      rq_wait_pos_spe_for_request(255, 204, 255, "1")
      rq_go_to("1")
      rq_wait("1")
      # end: URCap Program Node
      $ 2057 "Decap"
      $ 2058 "Action_Info≔'decapping'"
      global Action_Info="decapping"
      $ 2059 "Set GRP_3F_Enable=On"
      set_standard_digital_out(4, True)
      $ 2060 "Set GRP_3F_Decap=On"
      set_standard_digital_out(3, True)
      $ 2061 "Force"
      sleep(0.02)
      zero_ftsensor()
      force_mode(p[0.0,0.0,0.0,0.0,0.0,0.0], [0, 0, 1, 0, 0, 0], [0.0, 0.0, 1.0, 0.0, 0.0, 0.0], 2, [0.1, 0.1, 0.001, 0.3490658503988659, 0.3490658503988659, 0.3490658503988659])
      $ 2062 "check_decapping(offset=0.015, timeout=10, abort=CMD_Hold)" "noBreak"
      check_decapping(offset=0.015, timeout=10, abort=CMD_Hold)
      end_force_mode()
      stopl(5.0)
      $ 2063 "Set GRP_3F_Decap=Off"
      set_standard_digital_out(3, False)
      $ 2064 "Set GRP_3F_Enable=Off"
      set_standard_digital_out(4, False)
      $ 2065 "MoveL"
      $ 2066 "Waypoint_90" "breakAfter"
      movel(Waypoint_90_p, a=0.5, v=0.1, r=0.05)
      $ 2067 "MoveJ"
      $ 2068 "cap_dump_2" "breakAfter"
      movej(get_inverse_kin(cap_dump_2_p, qnear=cap_dump_2_q), a=0.5235987755982988, v=0.4363323129985824)
      # begin: URCap Program Node
      #   Source: Robotiq_Grippers, 3.17.0.105337, Robotiq Inc.
      #   Type: Gripper
      $ 2069 "Gripper Open (1)"
      if not(gripper_connected[0]):
        popup("Gripper 1 must be connected to run this program.", "No connection", False, True, True)
      end
      if not(rq_is_gripper_activated("1")):
        popup("Gripper 1 is not activated. Go to Installation tab > Gripper to activate it and run the program again.", "Not activated", False, True, True)
      end
      rq_set_pos_spd_for(0, 204, 255, "1")
      rq_wait_pos_spe_for_request(0, 204, 255, "1")
      rq_go_to("1")
      rq_wait("1")
      # end: URCap Program Node
      $ 2070 "MoveJ"
      $ 2071 "Waypoint_91" "breakAfter"
      movej(get_inverse_kin(Waypoint_91_p, qnear=Waypoint_91_q), a=0.5235987755982988, v=0.4363323129985824, r=0.036)
    elif (33 == switch_1):
      $ 2072 "Case 33"
      $ 2073 "Shake and liquid transfer"
      $ 2074 "MoveL"
      $ 2075 "Vial_liq_abov_1" "breakAfter"
      movel(Vial_liq_abov_1_p, a=0.5, v=0.1)
      $ 2076 "Vial_liq_pick_3" "breakAfter"
      movel(Vial_liq_pick_3_p, a=0.5, v=0.1)
      $ 2077 "Vial_liq_pick_4" "breakAfter"
      movel(Vial_liq_pick_4_p, a=0.5, v=0.1)
      # begin: URCap Program Node
      #   Source: Robotiq_Grippers, 3.17.0.105337, Robotiq Inc.
      #   Type: Gripper
      $ 2078 "Gripper Close (1)"
      if not(gripper_connected[0]):
        popup("Gripper 1 must be connected to run this program.", "No connection", False, True, True)
      end
      if not(rq_is_gripper_activated("1")):
        popup("Gripper 1 is not activated. Go to Installation tab > Gripper to activate it and run the program again.", "Not activated", False, True, True)
      end
      rq_set_pos_spd_for(255, 82, 71, "1")
      rq_wait_pos_spe_for_request(255, 82, 71, "1")
      rq_go_to("1")
      rq_wait("1")
      # end: URCap Program Node
      $ 2079 "Wait: 1.0"
      sleep(1.0)
      $ 2080 "Set GRP_3F_Open=On"
      set_standard_digital_out(5, True)
      $ 2081 "Wait: 0.5"
      sleep(0.5)
      $ 2082 "Vial_liq_abov_2" "breakAfter"
      movel(Vial_liq_abov_2_p, a=0.3, v=0.05, r=0.05)
      $ 2083 "MoveL"
      $ 2084 "Liquid_midway_1" "breakAfter"
      movel(Liquid_midway_1_p, a=0.5, v=0.1)
      $ 2085 "Loop 3 times"
      Loop_1 = 0
      while (Loop_1 < 3):
        $ 2086 "shake_3" "breakAfter"
        movel(shake_3_p, a=2.0, v=0.5)
        $ 2087 "shake_4" "breakAfter"
        movel(shake_4_p, a=2.0, v=0.5)
        Loop_1 = Loop_1 + 1
      end
      $ 2088 "drop_above_3" "breakAfter"
      movel(drop_above_3_p, a=0.5, v=0.1)
      $ 2089 "drop_above_4" "breakAfter"
      movel(drop_above_4_p, a=0.5, v=0.1)
      $ 2090 "liq_tran_3" "breakAfter"
      movel(liq_tran_3_p, a=0.5, v=0.05, r=0.008)
      $ 2091 "Wait: 1.0"
      sleep(1.0)
      $ 2092 "drop_above_5" "breakAfter"
      movel(drop_above_5_p, a=0.5, v=0.1)
      $ 2093 "Waypoint_92" "breakAfter"
      movel(Waypoint_92_p, a=0.5, v=0.1)
      $ 2094 "liq_tran_4" "breakAfter"
      movel(liq_tran_4_p, a=0.5, v=0.05)
      $ 2095 "Wait: 1.0"
      sleep(1.0)
      $ 2096 "drop_above_6" "breakAfter"
      movel(drop_above_6_p, a=0.5, v=0.1)
      $ 2097 "drop_above_7" "breakAfter"
      movel(drop_above_7_p, a=0.5, v=0.1)
      $ 2098 "Liquid_midway_2" "breakAfter"
      movel(Liquid_midway_2_p, a=0.5, v=0.1)
      $ 2099 "MoveL"
      $ 2100 "Vial_drop_abo_1" "breakAfter"
      movel(Vial_drop_abo_1_p, a=0.5, v=0.1)
      $ 2101 "Vial_liq_drop_1" "breakAfter"
      movel(Vial_liq_drop_1_p, a=0.5, v=0.1)
      # begin: URCap Program Node
      #   Source: Robotiq_Grippers, 3.17.0.105337, Robotiq Inc.
      #   Type: Gripper
      $ 2102 "Gripper Open (1)"
      if not(gripper_connected[0]):
        popup("Gripper 1 must be connected to run this program.", "No connection", False, True, True)
      end
      if not(rq_is_gripper_activated("1")):
        popup("Gripper 1 is not activated. Go to Installation tab > Gripper to activate it and run the program again.", "Not activated", False, True, True)
      end
      rq_set_pos_spd_for(0, 82, 71, "1")
      rq_wait_pos_spe_for_request(0, 82, 71, "1")
      rq_go_to("1")
      rq_wait("1")
      # end: URCap Program Node
      $ 2103 "Vial_drop_abo_2" "breakAfter"
      movel(Vial_drop_abo_2_p, a=0.5, v=0.1)
    elif (34 == switch_1):
      $ 2104 "Case 34"
      $ 2105 "Task≔'Dosing'"
      global Task="Dosing"
      $ 2106 "tilt_to_home()"
      tilt_to_home()
      $ 2107 "Powder dosing all"
      $ 2108 "tilt_angle_sent≔0.0"
      global tilt_angle_sent=0.0
      $ 2109 "send_target_info()"
      send_target_info()
      $ 2111 "prev_spat≔''"
      global prev_spat=""
      $ 2112 "spatula≔''"
      global spatula=""
      $ 2113 "scoop_status≔'normal'"
      global scoop_status="normal"
      $ 2114 "send_powder_info()"
      send_powder_info()
      $ 2115 "Set AO[0]=0.0"
      set_standard_analog_out(0, 0.0)
      $ 2116 "Wait: 0.2"
      sleep(0.2)
      $ 2117 "reach pots decapping pose"
      # begin: URCap Program Node
      #   Source: SensoPart VISOR Robotic, 2.0.6, SensoPart Industriesensorik GmbH
      #   Type: VISOR Robotic App
      $ 2123 "VISOR Easy Pick"
      def visorFuncEasyPick_4c19ec():
        # begin: URCap Program Node
        #   Source: SensoPart VISOR Robotic, 2.0.6, SensoPart Industriesensorik GmbH
        #   Type: Easy Pick Setup
        $ 2124 "# 1 Setup" "noBreak"
        local easyPickVisorId = 1
        local easyPickArmMounted = True
        local easyPickSetJob = True
        local easyPickJobName = "Weight_scale"
        local easyPickAtImgAcq = False
        local easyPickImgAcqPose = Trigger
        # end: URCap Program Node
        # begin: URCap Program Node
        #   Source: SensoPart VISOR Robotic, 2.0.6, SensoPart Industriesensorik GmbH
        #   Type: Process
        $ 2125 "Process" "noBreak"
        local easyPickObjTaken = False
        local easyPickTrigger = False
        local easyPickPoseIdx = 0
        local easyPickPose = p[0,0,0,0,0,0]
        def easyPickFuncTrigger(visorId, setJob, jobName, arm):
        if (setJob):
          visor_changeJob(visorId, jobName, 6000)
        end
        if (arm):
          visor_trigger(visorId, 6000, "arm")
        else:
          visor_trigger(visorId, 6000)
        end
        global easyPickParts_4=visor_partsFound(visorId)
        visor_easyPickUpdate(visorId, "parts", visor_partsFound(visorId))
        return visor_getPose3d(visorId, 0)
      end
      while (not easyPickObjTaken):
        easyPickTrigger = (easyPickCount_4 >= visor_partsFound(easyPickVisorId)) or (easyPickCount_4 > 9) or (not visor_easyPickCheckIdent("3d3650", easyPickVisorId))
        if (easyPickTrigger):
          easyPickCount_4 = 0
        end
        easyPickPoseIdx = easyPickCount_4
        easyPickPose = visor_getPose3d(easyPickVisorId, easyPickPoseIdx)
        visor_easyPickUpdate(easyPickVisorId, "counter", easyPickPoseIdx)
        # begin: URCap Program Node
        #   Source: SensoPart VISOR Robotic, 2.0.6, SensoPart Industriesensorik GmbH
        #   Type: Image Acquisition Pose
        $ 2126 "Image Acquisition Pose" "noBreak"
        if (easyPickTrigger):
          if (not easyPickAtImgAcq):
            movej(pose_trans(easyPickImgAcqPose,p[0.0000,0.0000,-0.0000,0.0000,0.0000,0.0000]),a=1.3963,v=1.0472,t=0.000000,r=0.000000)
            easyPickAtImgAcq = True
          end
          easyPickPose = easyPickFuncTrigger(easyPickVisorId, easyPickSetJob, easyPickJobName, easyPickArmMounted)
        end
        # end: URCap Program Node
        # begin: URCap Program Node
        #   Source: SensoPart VISOR Robotic, 2.0.6, SensoPart Industriesensorik GmbH
        #   Type: Object Detected
        $ 2127 "Object Detected" "noBreak"
        if (visor_partsFound(easyPickVisorId) > 0):
          $ 2128 "Open Gripper" "noBreak"
          $ 2129 "weight_value≔get_weight()" "noBreak"
          global weight_value=get_weight()
          $ 2130 "Wait: 0.5" "noBreak"
          sleep(0.5)
          $ 2131 "diff≔target_weight-weight_value" "noBreak"
          global diff=target_weight-weight_value
          $ 2132 "compute_level_percent(W_now, weight_value)" "noBreak"
          compute_level_percent(W_now, weight_value)
          $ 2133 "send_level_info()" "noBreak"
          send_level_info()
          $ 2134 "spatula≔select_spatula(Flowability, level, diff, bulk_density, mouth_d)" "noBreak"
          global spatula=select_spatula(Flowability, level, diff, bulk_density, mouth_d)
          $ 2135 "Wait: 0.2" "noBreak"
          sleep(0.2)
          $ 2136 "send_spatula_info()" "noBreak"
          send_spatula_info()
          $ 2137 "Pick spatula" "noBreak"
          $ 2138 "If spatula ≟ 'spatula_L'" "noBreak"
          if (spatula  ==  "spatula_L"):
            $ 2139 "MoveJ" "noBreak"
            $ 2140 "Spatula_otw" "noBreak"
            movej(get_inverse_kin(Spatula_otw_p, qnear=Spatula_otw_q), a=1.3962634015954636, v=1.0471975511965976)
            $ 2141 "pick_spat_L_abv" "noBreak"
            movej(get_inverse_kin(pick_spat_L_abv_p, qnear=pick_spat_L_abv_q), a=1.3962634015954636, v=1.0471975511965976)
            $ 2142 "MoveL" "noBreak"
            $ 2143 "spat_L_pick" "noBreak"
            movel(spat_L_pick_p, a=1.2, v=0.25)
            # begin: URCap Program Node
            #   Source: Robotiq_Grippers, 3.17.0.105337, Robotiq Inc.
            #   Type: Gripper
            $ 2144 "Gripper Close (1)" "noBreak"
            if not(gripper_connected[0]):
              popup("Gripper 1 must be connected to run this program.", "No connection", False, True, True)
            end
            if not(rq_is_gripper_activated("1")):
              popup("Gripper 1 is not activated. Go to Installation tab > Gripper to activate it and run the program again.", "Not activated", False, True, True)
            end
            rq_set_pos_spd_for(255, 0, 77, "1")
            rq_wait_pos_spe_for_request(255, 0, 77, "1")
            rq_go_to("1")
            rq_wait("1")
            # end: URCap Program Node
            $ 2145 "spat_L_lift" "noBreak"
            movel(spat_L_lift_p, a=1.2, v=0.25, r=0.01)
            $ 2146 "spat_L_side" "noBreak"
            movel(spat_L_side_p, a=1.2, v=0.25, r=0.01)
            $ 2147 "spat_L_up" "noBreak"
            movel(spat_L_up_p, a=1.2, v=0.25, r=0.05)
            $ 2148 "MoveJ" "noBreak"
            $ 2149 "Spatula_otw" "noBreak"
            movej(get_inverse_kin(Spatula_otw_p, qnear=Spatula_otw_q), a=1.3962634015954636, v=1.0471975511965976)
          else:
            $ 2150 "ElseIf spatula ≟'spatula_M'" "noBreak"
            if (spatula  == "spatula_M"):
              $ 2151 "MoveJ" "noBreak"
              $ 2152 "Spatula_otw" "noBreak"
              movej(get_inverse_kin(Spatula_otw_p, qnear=Spatula_otw_q), a=1.3962634015954636, v=1.0471975511965976)
              $ 2153 "spat_M_up" "noBreak"
              movej(get_inverse_kin(spat_M_up_p, qnear=spat_M_up_q), a=1.3962634015954636, v=1.0471975511965976, r=0.05)
              $ 2154 "MoveL" "noBreak"
              $ 2155 "spat_M_pick" "noBreak"
              movel(spat_M_pick_p, a=1.2, v=0.25)
              # begin: URCap Program Node
              #   Source: Robotiq_Grippers, 3.17.0.105337, Robotiq Inc.
              #   Type: Gripper
              $ 2156 "Gripper Close (1)" "noBreak"
              if not(gripper_connected[0]):
                popup("Gripper 1 must be connected to run this program.", "No connection", False, True, True)
              end
              if not(rq_is_gripper_activated("1")):
                popup("Gripper 1 is not activated. Go to Installation tab > Gripper to activate it and run the program again.", "Not activated", False, True, True)
              end
              rq_set_pos_spd_for(255, 0, 77, "1")
              rq_wait_pos_spe_for_request(255, 0, 77, "1")
              rq_go_to("1")
              rq_wait("1")
              # end: URCap Program Node
              $ 2157 "spat_M_up" "noBreak"
              movel(spat_M_up_p, a=1.2, v=0.25, r=0.05)
              $ 2158 "Spatula_otw" "noBreak"
              movel(Spatula_otw_p, a=1.2, v=0.25)
              $ 2159 "switch_spat_M≔ False " "noBreak"
              global switch_spat_M=  False
            else:
              $ 2160 "ElseIf spatula≟'spatula_S'" "noBreak"
              if (spatula == "spatula_S"):
                $ 2161 "MoveJ" "noBreak"
                $ 2162 "Spatula_otw" "noBreak"
                movej(get_inverse_kin(Spatula_otw_p, qnear=Spatula_otw_q), a=1.3962634015954636, v=1.0471975511965976)
                $ 2163 "spat_S_Up_7" "noBreak"
                movej(get_inverse_kin(spat_S_Up_7_p, qnear=spat_S_Up_7_q), a=1.3962634015954636, v=1.0471975511965976, r=0.05)
                $ 2164 "MoveL" "noBreak"
                $ 2165 "spat_S_Pick_4" "noBreak"
                movel(spat_S_Pick_4_p, a=1.2, v=0.25)
                # begin: URCap Program Node
                #   Source: Robotiq_Grippers, 3.17.0.105337, Robotiq Inc.
                #   Type: Gripper
                $ 2166 "Gripper Close (1)" "noBreak"
                if not(gripper_connected[0]):
                  popup("Gripper 1 must be connected to run this program.", "No connection", False, True, True)
                end
                if not(rq_is_gripper_activated("1")):
                  popup("Gripper 1 is not activated. Go to Installation tab > Gripper to activate it and run the program again.", "Not activated", False, True, True)
                end
                rq_set_pos_spd_for(255, 0, 77, "1")
                rq_wait_pos_spe_for_request(255, 0, 77, "1")
                rq_go_to("1")
                rq_wait("1")
                # end: URCap Program Node
                $ 2167 "spat_S_Up_8" "noBreak"
                movel(spat_S_Up_8_p, a=1.2, v=0.25, r=0.05)
                $ 2168 "Spatula_otw" "noBreak"
                movel(Spatula_otw_p, a=1.2, v=0.25)
                $ 2169 "switch_spat_S≔ False " "noBreak"
                global switch_spat_S=  False
              else:
                $ 2170 "ElseIf spatula≟'spatula_flat_M'" "noBreak"
                if (spatula == "spatula_flat_M"):
                  $ 2171 "MoveJ" "noBreak"
                  $ 2172 "Spatula_otw" "noBreak"
                  movej(get_inverse_kin(Spatula_otw_p, qnear=Spatula_otw_q), a=1.3962634015954636, v=1.0471975511965976)
                  $ 2173 "spat_flatM_up" "noBreak"
                  movej(get_inverse_kin(spat_flatM_up_p, qnear=spat_flatM_up_q), a=1.3962634015954636, v=1.0471975511965976, r=0.05)
                  $ 2174 "MoveL" "noBreak"
                  $ 2175 "spat_flatM_pick" "noBreak"
                  movel(spat_flatM_pick_p, a=1.2, v=0.25)
                  # begin: URCap Program Node
                  #   Source: Robotiq_Grippers, 3.17.0.105337, Robotiq Inc.
                  #   Type: Gripper
                  $ 2176 "Gripper Close (1)" "noBreak"
                  if not(gripper_connected[0]):
                    popup("Gripper 1 must be connected to run this program.", "No connection", False, True, True)
                  end
                  if not(rq_is_gripper_activated("1")):
                    popup("Gripper 1 is not activated. Go to Installation tab > Gripper to activate it and run the program again.", "Not activated", False, True, True)
                  end
                  rq_set_pos_spd_for(255, 0, 77, "1")
                  rq_wait_pos_spe_for_request(255, 0, 77, "1")
                  rq_go_to("1")
                  rq_wait("1")
                  # end: URCap Program Node
                  $ 2177 "spat_flatM_up" "noBreak"
                  movel(spat_flatM_up_p, a=1.2, v=0.25, r=0.05)
                  $ 2178 "Spatula_otw" "noBreak"
                  movel(Spatula_otw_p, a=1.2, v=0.25)
                  $ 2179 "switch_spat_F_M≔ False " "noBreak"
                  global switch_spat_F_M=  False
                else:
                  $ 2180 "ElseIf spatula≟'spatula_flat_S'" "noBreak"
                  if (spatula == "spatula_flat_S"):
                    $ 2181 "MoveJ" "noBreak"
                    $ 2182 "Spatula_otw" "noBreak"
                    movej(get_inverse_kin(Spatula_otw_p, qnear=Spatula_otw_q), a=1.3962634015954636, v=1.0471975511965976)
                    $ 2183 "spat_flatS_up" "noBreak"
                    movej(get_inverse_kin(spat_flatS_up_p, qnear=spat_flatS_up_q), a=1.3962634015954636, v=1.0471975511965976, r=0.05)
                    $ 2184 "MoveL" "noBreak"
                    $ 2185 "spat_flatS_pick" "noBreak"
                    movel(spat_flatS_pick_p, a=1.2, v=0.25)
                    # begin: URCap Program Node
                    #   Source: Robotiq_Grippers, 3.17.0.105337, Robotiq Inc.
                    #   Type: Gripper
                    $ 2186 "Gripper Close (1)" "noBreak"
                    if not(gripper_connected[0]):
                      popup("Gripper 1 must be connected to run this program.", "No connection", False, True, True)
                    end
                    if not(rq_is_gripper_activated("1")):
                      popup("Gripper 1 is not activated. Go to Installation tab > Gripper to activate it and run the program again.", "Not activated", False, True, True)
                    end
                    rq_set_pos_spd_for(255, 0, 77, "1")
                    rq_wait_pos_spe_for_request(255, 0, 77, "1")
                    rq_go_to("1")
                    rq_wait("1")
                    # end: URCap Program Node
                    $ 2187 "spat_flatS_up" "noBreak"
                    movel(spat_flatS_up_p, a=1.2, v=0.25, r=0.05)
                    $ 2188 "Spatula_otw" "noBreak"
                    movel(Spatula_otw_p, a=1.2, v=0.25)
                    $ 2189 "switch_spat_F_S≔ False " "noBreak"
                    global switch_spat_F_S=  False
                  end
                end
              end
            end
          end
          $ 2190 "Action_Info≔'Scooping'" "noBreak"
          global Action_Info="Scooping"
          $ 2191 "auto_tilt_and_scoop(W_now, target_weight, weight_value)" "noBreak"
          auto_tilt_and_scoop(W_now, target_weight, weight_value)
          $ 2192 "Action_Info≔'Dosing'" "noBreak"
          global Action_Info="Dosing"
          # begin: URCap Program Node
          #   Source: SensoPart VISOR Robotic, 2.0.6, SensoPart Industriesensorik GmbH
          #   Type: Approach Pose
          $ 2193 "Approach Pose" "noBreak"
          movej(pose_trans(easyPickPose,p[0.0000,0.0000,-0.0000,0.0000,0.0000,0.0000]),a=0.2618,v=0.1745,t=0.000000,r=0.000000)
          # end: URCap Program Node
          # begin: URCap Program Node
          #   Source: SensoPart VISOR Robotic, 2.0.6, SensoPart Industriesensorik GmbH
          #   Type: Target Pose
          $ 2194 "Target Pose" "noBreak"
          movel(pose_trans(easyPickPose,p[0.0000,0.0000,-0.0000,0.0000,0.0000,0.0000]),a=0.0500,v=0.0200,t=0.000000,r=0.000000)
          # end: URCap Program Node
          $ 2195 "Close Gripper" "noBreak"
          $ 2196 "current_p≔get_actual_tcp_pose()" "noBreak"
          global current_p= get_actual_tcp_pose ()
          $ 2197 "dispense_pos≔pose_trans(current_p,p[0,0,0,0,-deg2rad(spatula_ry),0])" "noBreak"
          global dispense_pos=pose_trans(current_p,p[0,0,0,0,-deg2rad(spatula_ry),0])
          $ 2198 "Loop weight_value≤target_weight and delta_count≤3" "noBreak"
          thread Thread_while_2198():
            while (True):
              $ 2199 "MoveL" "noBreak"
              $ 2200 "dispense_pos" "noBreak"
              movel(dispense_pos, a=0.2, v=0.1)
              $ 2201 "log_weight()" "noBreak"
              log_weight()
              $ 2203 "CCW_full_Rotate()" "noBreak"
              CCW_full_Rotate()
              $ 2204 "Start_thread≔ True " "noBreak"
              global Start_thread=  True
              $ 2205 "vib_thread≔ True " "noBreak"
              global vib_thread=  True
              $ 2206 "Wait: 0.5" "noBreak"
              sleep(0.5)
              $ 2207 "If diff ≥(target_g*1.2)" "noBreak"
              if (diff  >= (target_g*1.2)):
                $ 2208 "tilt_pose≔pose_trans(get_actual_tcp_pose(), p[0, 0, 0, 0, 0, 2.0])" "noBreak"
                global tilt_pose=pose_trans(get_actual_tcp_pose(), p[0, 0, 0, 0, 0, 2.0])
                $ 2209 "movel(tilt_pose, a=0.5, v=0.5, r=0.00001)" "noBreak"
                movel(tilt_pose, a=0.5, v=0.5, r=0.00001)
              else:
                $ 2210 "Else" "noBreak"
                $ 2211 "Loop weight_value≤(target_weight-0.00) and tilt_angle≥(-1.999) and tilt_angle≤0.5" "noBreak"
                thread Thread_while_2211():
                  while (True):
                    $ 2212 "current_error≔target_weight-weight_value" "noBreak"
                    global current_error=target_weight-weight_value
                    $ 2213 "Integral_error≔Integral_error+current_error*dt" "noBreak"
                    global Integral_error=Integral_error+current_error*dt
                    $ 2214 "derivative≔(current_error-previous_error)/dt" "noBreak"
                    global derivative=(current_error-previous_error)/dt
                    $ 2215 "tilt_increment≔(kp*current_error)+(ki*Integral_error)+(kd*derivative)" "noBreak"
                    global tilt_increment=(kp*current_error)+(ki*Integral_error)+(kd*derivative)
                    $ 2216 "current_pose≔get_actual_tcp_pose()" "noBreak"
                    global current_pose= get_actual_tcp_pose ()
                    $ 2217 "tilt_angle≔current_pose[5]" "noBreak"
                    global tilt_angle=current_pose[5]
                    $ 2218 "tilt_pose≔pose_trans(current_pose, p[0, 0, 0, 0, 0, tilt_increment])" "noBreak"
                    global tilt_pose=pose_trans(current_pose, p[0, 0, 0, 0, 0, tilt_increment])
                    $ 2219 "movel(tilt_pose, a=0.1, v=0.1, r=0.00001)" "noBreak"
                    movel(tilt_pose, a=0.1, v=0.1, r=0.00001)
                    $ 2220 "previous_error≔current_error" "noBreak"
                    global previous_error=current_error
                  end
                end
                if (weight_value <= (target_weight-0.00)  and  tilt_angle >= (-1.999)  and  tilt_angle <= 0.5):
                  global thread_handler_2211=run Thread_while_2211()
                  while (weight_value <= (target_weight-0.00)  and  tilt_angle >= (-1.999)  and  tilt_angle <= 0.5):
                    sync()
                  end
                  kill thread_handler_2211
                end
              end
              $ 2221 "weight_value≔get_weight()" "noBreak"
              global weight_value=get_weight()
              $ 2222 "tilt_angle≔-1" "noBreak"
              global tilt_angle=-1
              $ 2223 "Wait: 0.5" "noBreak"
              sleep(0.5)
              $ 2224 "Start_thread≔ False " "noBreak"
              global Start_thread=  False
              $ 2225 "vib_thread≔ False " "noBreak"
              global vib_thread=  False
              $ 2226 "dispense_pos" "noBreak"
              movel(dispense_pos, a=1.2, v=0.25)
              $ 2227 "compute_level_percent(W_now, weight_value)" "noBreak"
              compute_level_percent(W_now, weight_value)
              $ 2228 "If delta<0.01" "noBreak"
              if (delta<0.01):
                $ 2229 "delta_count≔delta_count+1" "noBreak"
                global delta_count=delta_count+1
              else:
                $ 2230 "Else" "noBreak"
                $ 2231 "delta_count≔0" "noBreak"
                global delta_count=0
              end
              $ 2232 "prev_spat≔spatula" "noBreak"
              global prev_spat=spatula
              $ 2233 "Wait: 0.2" "noBreak"
              sleep(0.2)
              $ 2234 "spatula≔select_spatula(Flowability, level, diff, bulk_density, mouth_d)" "noBreak"
              global spatula=select_spatula(Flowability, level, diff, bulk_density, mouth_d)
              $ 2235 "Wait: 1.0" "noBreak"
              sleep(1.0)
              $ 2236 "send_level_info()" "noBreak"
              send_level_info()
              $ 2237 "send_spatula_info()" "noBreak"
              send_spatula_info()
              $ 2238 "Integral_error≔0" "noBreak"
              global Integral_error=0
              $ 2239 "current_error≔0" "noBreak"
              global current_error=0
              $ 2240 "previous_error≔0" "noBreak"
              global previous_error=0
              $ 2241 "Set AO[0]=0.0" "noBreak"
              set_standard_analog_out(0, 0.0)
              $ 2242 "Wait: 0.5" "noBreak"
              sleep(0.5)
              $ 2243 "swtich spatula" "noBreak"
              $ 2244 "If spatula ≟ 'spatula_M' and switch_spat_M≟ True " "noBreak"
              if (spatula  ==  "spatula_M"  and  switch_spat_M ==   True  ):
                $ 2245 "MoveJ" "noBreak"
                $ 2246 "Spatula_otw" "noBreak"
                movej(get_inverse_kin(Spatula_otw_p, qnear=Spatula_otw_q), a=1.3962634015954636, v=1.0471975511965976)
                $ 2247 "spat_L_up" "noBreak"
                movej(get_inverse_kin(spat_L_up_p, qnear=spat_L_up_q), a=1.3962634015954636, v=1.0471975511965976)
                $ 2248 "MoveL" "noBreak"
                $ 2249 "spat_L_side" "noBreak"
                movel(spat_L_side_p, a=1.2, v=0.25)
                $ 2250 "spat_L_lift" "noBreak"
                movel(spat_L_lift_p, a=1.2, v=0.25)
                $ 2251 "spat_L_pick" "noBreak"
                movel(spat_L_pick_p, a=0.2, v=0.1)
                # begin: URCap Program Node
                #   Source: Robotiq_Grippers, 3.17.0.105337, Robotiq Inc.
                #   Type: Gripper
                $ 2252 "Gripper Open (1)" "noBreak"
                if not(gripper_connected[0]):
                  popup("Gripper 1 must be connected to run this program.", "No connection", False, True, True)
                end
                if not(rq_is_gripper_activated("1")):
                  popup("Gripper 1 is not activated. Go to Installation tab > Gripper to activate it and run the program again.", "Not activated", False, True, True)
                end
                rq_set_pos_spd_for(0, 255, 77, "1")
                rq_wait_pos_spe_for_request(0, 255, 77, "1")
                rq_go_to("1")
                rq_wait("1")
                # end: URCap Program Node
                $ 2253 "spat_M_pick" "noBreak"
                movel(spat_M_pick_p, a=1.2, v=0.25)
                # begin: URCap Program Node
                #   Source: Robotiq_Grippers, 3.17.0.105337, Robotiq Inc.
                #   Type: Gripper
                $ 2254 "Gripper Close (1)" "noBreak"
                if not(gripper_connected[0]):
                  popup("Gripper 1 must be connected to run this program.", "No connection", False, True, True)
                end
                if not(rq_is_gripper_activated("1")):
                  popup("Gripper 1 is not activated. Go to Installation tab > Gripper to activate it and run the program again.", "Not activated", False, True, True)
                end
                rq_set_pos_spd_for(255, 0, 77, "1")
                rq_wait_pos_spe_for_request(255, 0, 77, "1")
                rq_go_to("1")
                rq_wait("1")
                # end: URCap Program Node
                $ 2255 "spat_M_up" "noBreak"
                movel(spat_M_up_p, a=1.2, v=0.25)
                $ 2256 "Spatula_otw" "noBreak"
                movel(Spatula_otw_p, a=1.2, v=0.25)
                $ 2257 "switch_spat_M≔ False " "noBreak"
                global switch_spat_M=  False
                $ 2258 "correction_reset()" "noBreak"
                correction_reset()
              else:
                $ 2259 "ElseIf spatula ≟ 'spatula_S' and switch_spat_S ≟ True and prev_spat≟'spatula_M'" "noBreak"
                if (spatula  ==  "spatula_S" and switch_spat_S  ==   True  and prev_spat == "spatula_M"):
                  $ 2260 "MoveL" "noBreak"
                  $ 2261 "Spatula_otw" "noBreak"
                  movel(Spatula_otw_p, a=1.2, v=0.25)
                  $ 2262 "spat_M_up" "noBreak"
                  movel(spat_M_up_p, a=1.2, v=0.25)
                  $ 2263 "spat_M_pick" "noBreak"
                  movel(spat_M_pick_p, a=0.2, v=0.1)
                  # begin: URCap Program Node
                  #   Source: Robotiq_Grippers, 3.17.0.105337, Robotiq Inc.
                  #   Type: Gripper
                  $ 2264 "Gripper Open (1)" "noBreak"
                  if not(gripper_connected[0]):
                    popup("Gripper 1 must be connected to run this program.", "No connection", False, True, True)
                  end
                  if not(rq_is_gripper_activated("1")):
                    popup("Gripper 1 is not activated. Go to Installation tab > Gripper to activate it and run the program again.", "Not activated", False, True, True)
                  end
                  rq_set_pos_spd_for(0, 255, 77, "1")
                  rq_wait_pos_spe_for_request(0, 255, 77, "1")
                  rq_go_to("1")
                  rq_wait("1")
                  # end: URCap Program Node
                  $ 2265 "spat_S_pick" "noBreak"
                  movel(spat_S_pick_p, a=1.2, v=0.25)
                  # begin: URCap Program Node
                  #   Source: Robotiq_Grippers, 3.17.0.105337, Robotiq Inc.
                  #   Type: Gripper
                  $ 2266 "Gripper Close (1)" "noBreak"
                  if not(gripper_connected[0]):
                    popup("Gripper 1 must be connected to run this program.", "No connection", False, True, True)
                  end
                  if not(rq_is_gripper_activated("1")):
                    popup("Gripper 1 is not activated. Go to Installation tab > Gripper to activate it and run the program again.", "Not activated", False, True, True)
                  end
                  rq_set_pos_spd_for(255, 0, 77, "1")
                  rq_wait_pos_spe_for_request(255, 0, 77, "1")
                  rq_go_to("1")
                  rq_wait("1")
                  # end: URCap Program Node
                  $ 2267 "spat_S_up" "noBreak"
                  movel(spat_S_up_p, a=1.2, v=0.25)
                  $ 2268 "Spatula_otw" "noBreak"
                  movel(Spatula_otw_p, a=1.2, v=0.25)
                  $ 2269 "switch_spat_S≔ False " "noBreak"
                  global switch_spat_S=  False
                  $ 2270 "correction_reset()" "noBreak"
                  correction_reset()
                else:
                  $ 2271 "ElseIf spatula≟'spatula_S' and switch_spat_S≟ True  and prev_spat≟'spatula_L'" "noBreak"
                  if (spatula == "spatula_S" and switch_spat_S ==   True    and  prev_spat == "spatula_L"):
                    $ 2272 "MoveJ" "noBreak"
                    $ 2273 "Spatula_otw" "noBreak"
                    movej(get_inverse_kin(Spatula_otw_p, qnear=Spatula_otw_q), a=1.3962634015954636, v=1.0471975511965976)
                    $ 2274 "spat_L_up" "noBreak"
                    movej(get_inverse_kin(spat_L_up_p, qnear=spat_L_up_q), a=1.3962634015954636, v=1.0471975511965976)
                    $ 2275 "MoveL" "noBreak"
                    $ 2276 "spat_L_side" "noBreak"
                    movel(spat_L_side_p, a=1.2, v=0.25)
                    $ 2277 "spat_L_lift" "noBreak"
                    movel(spat_L_lift_p, a=1.2, v=0.25)
                    $ 2278 "spat_L_pick" "noBreak"
                    movel(spat_L_pick_p, a=0.2, v=0.1)
                    # begin: URCap Program Node
                    #   Source: Robotiq_Grippers, 3.17.0.105337, Robotiq Inc.
                    #   Type: Gripper
                    $ 2279 "Gripper Open (1)" "noBreak"
                    if not(gripper_connected[0]):
                      popup("Gripper 1 must be connected to run this program.", "No connection", False, True, True)
                    end
                    if not(rq_is_gripper_activated("1")):
                      popup("Gripper 1 is not activated. Go to Installation tab > Gripper to activate it and run the program again.", "Not activated", False, True, True)
                    end
                    rq_set_pos_spd_for(0, 255, 77, "1")
                    rq_wait_pos_spe_for_request(0, 255, 77, "1")
                    rq_go_to("1")
                    rq_wait("1")
                    # end: URCap Program Node
                    $ 2280 "spat_S_pick" "noBreak"
                    movel(spat_S_pick_p, a=1.2, v=0.25)
                    # begin: URCap Program Node
                    #   Source: Robotiq_Grippers, 3.17.0.105337, Robotiq Inc.
                    #   Type: Gripper
                    $ 2281 "Gripper Close (1)" "noBreak"
                    if not(gripper_connected[0]):
                      popup("Gripper 1 must be connected to run this program.", "No connection", False, True, True)
                    end
                    if not(rq_is_gripper_activated("1")):
                      popup("Gripper 1 is not activated. Go to Installation tab > Gripper to activate it and run the program again.", "Not activated", False, True, True)
                    end
                    rq_set_pos_spd_for(255, 0, 77, "1")
                    rq_wait_pos_spe_for_request(255, 0, 77, "1")
                    rq_go_to("1")
                    rq_wait("1")
                    # end: URCap Program Node
                    $ 2282 "spat_S_up" "noBreak"
                    movel(spat_S_up_p, a=1.2, v=0.25)
                    $ 2283 "Spatula_otw" "noBreak"
                    movel(Spatula_otw_p, a=1.2, v=0.25)
                    $ 2284 "switch_spat_S≔ False " "noBreak"
                    global switch_spat_S=  False
                    $ 2285 "correction_reset()" "noBreak"
                    correction_reset()
                  else:
                    $ 2286 "ElseIf spatula≟'spatula_flat_S'  and switch_spat_F_S ≟ True " "noBreak"
                    if (spatula == "spatula_flat_S"   and  switch_spat_F_S  ==   True  ):
                      $ 2287 "MoveL" "noBreak"
                      $ 2288 "Spatula_otw" "noBreak"
                      movel(Spatula_otw_p, a=1.2, v=0.25)
                      $ 2289 "spat_flatM_up" "noBreak"
                      movel(spat_flatM_up_p, a=1.2, v=0.25)
                      $ 2290 "spat_flatM_pick" "noBreak"
                      movel(spat_flatM_pick_p, a=0.2, v=0.1)
                      # begin: URCap Program Node
                      #   Source: Robotiq_Grippers, 3.17.0.105337, Robotiq Inc.
                      #   Type: Gripper
                      $ 2291 "Gripper Open (1)" "noBreak"
                      if not(gripper_connected[0]):
                        popup("Gripper 1 must be connected to run this program.", "No connection", False, True, True)
                      end
                      if not(rq_is_gripper_activated("1")):
                        popup("Gripper 1 is not activated. Go to Installation tab > Gripper to activate it and run the program again.", "Not activated", False, True, True)
                      end
                      rq_set_pos_spd_for(0, 255, 74, "1")
                      rq_wait_pos_spe_for_request(0, 255, 74, "1")
                      rq_go_to("1")
                      rq_wait("1")
                      # end: URCap Program Node
                      $ 2292 "spat_flatS_pick" "noBreak"
                      movel(spat_flatS_pick_p, a=1.2, v=0.25)
                      # begin: URCap Program Node
                      #   Source: Robotiq_Grippers, 3.17.0.105337, Robotiq Inc.
                      #   Type: Gripper
                      $ 2293 "Gripper Close (1)" "noBreak"
                      if not(gripper_connected[0]):
                        popup("Gripper 1 must be connected to run this program.", "No connection", False, True, True)
                      end
                      if not(rq_is_gripper_activated("1")):
                        popup("Gripper 1 is not activated. Go to Installation tab > Gripper to activate it and run the program again.", "Not activated", False, True, True)
                      end
                      rq_set_pos_spd_for(255, 0, 77, "1")
                      rq_wait_pos_spe_for_request(255, 0, 77, "1")
                      rq_go_to("1")
                      rq_wait("1")
                      # end: URCap Program Node
                      $ 2294 "spat_flatS_up" "noBreak"
                      movel(spat_flatS_up_p, a=1.2, v=0.25)
                      $ 2295 "Spatula_otw" "noBreak"
                      movel(Spatula_otw_p, a=1.2, v=0.25)
                      $ 2296 "switch_spat_F_S≔ False " "noBreak"
                      global switch_spat_F_S=  False
                      $ 2297 "correction_reset()" "noBreak"
                      correction_reset()
                    end
                  end
                end
              end
              $ 2298 "tilt(level)" "noBreak"
              tilt(level)
              $ 2299 "Action_Info≔'Scooping'" "noBreak"
              global Action_Info="Scooping"
              $ 2300 "auto_tilt_and_scoop(W_now, target_weight, weight_value)" "noBreak"
              auto_tilt_and_scoop(W_now, target_weight, weight_value)
              $ 2301 "Action_Info≔'Dosing'" "noBreak"
              global Action_Info="Dosing"
            end
          end
          if (weight_value <= target_weight and delta_count <= 3):
            global thread_handler_2198=run Thread_while_2198()
            while (weight_value <= target_weight and delta_count <= 3):
              sync()
            end
            kill thread_handler_2198
          end
          $ 2302 "Start_thread≔ False " "noBreak"
          global Start_thread=  False
          $ 2303 "vib_thread≔ False " "noBreak"
          global vib_thread=  False
          # begin: URCap Program Node
          #   Source: SensoPart VISOR Robotic, 2.0.6, SensoPart Industriesensorik GmbH
          #   Type: Exit Pose
          $ 2304 "Exit Pose" "noBreak"
          movel(pose_trans(easyPickPose,p[0.0000,0.0000,-0.0000,0.0000,0.0000,0.0000]),a=0.5000,v=0.2500,t=0.000000,r=0.000000)
          # end: URCap Program Node
          easyPickObjTaken = True
        end
        # end: URCap Program Node
        # begin: URCap Program Node
        #   Source: SensoPart VISOR Robotic, 2.0.6, SensoPart Industriesensorik GmbH
        #   Type: No Object Detected
        $ 2305 "No Object Detected" "noBreak"
        if (visor_partsFound(easyPickVisorId) < 1):
          $ 2306 "Popup: No weigh scale detected" "noBreak"
          popup("No weigh scale detected", "Message", False, False, blocking=True)
          else:
        end
        # end: URCap Program Node
      end
      easyPickCount_4 = easyPickCount_4 + 1
      visor_easyPickUpdate(easyPickVisorId, "counter", easyPickCount_4)
      visor_easyPickSetIdent("3d3650", easyPickVisorId)
      # end: URCap Program Node
    end
    visorFuncEasyPick_4c19ec()
    # end: URCap Program Node
    $ 2307 "MoveL"
    $ 2308 "dispense_pos" "breakAfter"
    movel(dispense_pos, a=0.2, v=0.1)
    $ 2309 "after_scoop()"
    after_scoop()
    $ 2310 "Place spatula back to the rack"
    $ 2311 "If spatula ≟ 'spatula_L'"
    if (spatula  ==  "spatula_L"):
      $ 2312 "MoveJ"
      $ 2313 "Spatula_otw" "breakAfter"
      movej(get_inverse_kin(Spatula_otw_p, qnear=Spatula_otw_q), a=1.3962634015954636, v=1.0471975511965976)
      $ 2314 "MoveL"
      $ 2315 "spat_L_up" "breakAfter"
      movel(spat_L_up_p, a=1.2, v=0.25, r=0.05)
      $ 2316 "spat_L_side" "breakAfter"
      movel(spat_L_side_p, a=1.2, v=0.25, r=0.01)
      $ 2317 "spat_L_lift" "breakAfter"
      movel(spat_L_lift_p, a=1.2, v=0.25, r=0.01)
      $ 2318 "spat_L_pick" "breakAfter"
      movel(spat_L_pick_p, a=0.2, v=0.1)
      # begin: URCap Program Node
      #   Source: Robotiq_Grippers, 3.17.0.105337, Robotiq Inc.
      #   Type: Gripper
      $ 2319 "Gripper Open (1)"
      if not(gripper_connected[0]):
        popup("Gripper 1 must be connected to run this program.", "No connection", False, True, True)
      end
      if not(rq_is_gripper_activated("1")):
        popup("Gripper 1 is not activated. Go to Installation tab > Gripper to activate it and run the program again.", "Not activated", False, True, True)
      end
      rq_set_pos_spd_for(0, 128, 128, "1")
      rq_wait_pos_spe_for_request(0, 128, 128, "1")
      rq_go_to("1")
      rq_wait("1")
      # end: URCap Program Node
      $ 2320 "MoveJ"
      $ 2321 "pick_spat_L_abv" "breakAfter"
      movej(get_inverse_kin(pick_spat_L_abv_p, qnear=pick_spat_L_abv_q), a=1.3962634015954636, v=1.0471975511965976)
      $ 2322 "Spatula_otw" "breakAfter"
      movej(get_inverse_kin(Spatula_otw_p, qnear=Spatula_otw_q), a=1.3962634015954636, v=1.0471975511965976)
    else:
      $ 2323 "ElseIf spatula ≟'spatula_M'"
      if (spatula  == "spatula_M"):
        $ 2324 "MoveJ"
        $ 2325 "Spatula_otw" "breakAfter"
        movej(get_inverse_kin(Spatula_otw_p, qnear=Spatula_otw_q), a=1.3962634015954636, v=1.0471975511965976)
        $ 2326 "spat_M_up" "breakAfter"
        movej(get_inverse_kin(spat_M_up_p, qnear=spat_M_up_q), a=1.3962634015954636, v=1.0471975511965976, r=0.05)
        $ 2327 "MoveL"
        $ 2328 "spat_M_pick" "breakAfter"
        movel(spat_M_pick_p, a=0.2, v=0.1)
        # begin: URCap Program Node
        #   Source: Robotiq_Grippers, 3.17.0.105337, Robotiq Inc.
        #   Type: Gripper
        $ 2329 "Gripper Open (1)"
        if not(gripper_connected[0]):
          popup("Gripper 1 must be connected to run this program.", "No connection", False, True, True)
        end
        if not(rq_is_gripper_activated("1")):
          popup("Gripper 1 is not activated. Go to Installation tab > Gripper to activate it and run the program again.", "Not activated", False, True, True)
        end
        rq_set_pos_spd_for(0, 128, 128, "1")
        rq_wait_pos_spe_for_request(0, 128, 128, "1")
        rq_go_to("1")
        rq_wait("1")
        # end: URCap Program Node
        $ 2330 "spat_M_up" "breakAfter"
        movel(spat_M_up_p, a=1.2, v=0.25, r=0.05)
        $ 2331 "Spatula_otw" "breakAfter"
        movel(Spatula_otw_p, a=1.2, v=0.25)
        $ 2332 "switch_spat_M≔ False "
        global switch_spat_M=  False
      else:
        $ 2333 "ElseIf spatula≟'spatula_S'"
        if (spatula == "spatula_S"):
          $ 2334 "MoveJ"
          $ 2335 "Spatula_otw" "breakAfter"
          movej(get_inverse_kin(Spatula_otw_p, qnear=Spatula_otw_q), a=1.3962634015954636, v=1.0471975511965976)
          $ 2336 "spat_S_Up_7" "breakAfter"
          movej(get_inverse_kin(spat_S_Up_7_p, qnear=spat_S_Up_7_q), a=1.3962634015954636, v=1.0471975511965976, r=0.05)
          $ 2337 "MoveL"
          $ 2338 "spat_S_Pick_4" "breakAfter"
          movel(spat_S_Pick_4_p, a=0.2, v=0.1)
          # begin: URCap Program Node
          #   Source: Robotiq_Grippers, 3.17.0.105337, Robotiq Inc.
          #   Type: Gripper
          $ 2339 "Gripper Open (1)"
          if not(gripper_connected[0]):
            popup("Gripper 1 must be connected to run this program.", "No connection", False, True, True)
          end
          if not(rq_is_gripper_activated("1")):
            popup("Gripper 1 is not activated. Go to Installation tab > Gripper to activate it and run the program again.", "Not activated", False, True, True)
          end
          rq_set_pos_spd_for(0, 255, 51, "1")
          rq_wait_pos_spe_for_request(0, 255, 51, "1")
          rq_go_to("1")
          rq_wait("1")
          # end: URCap Program Node
          $ 2340 "spat_S_Up_8" "breakAfter"
          movel(spat_S_Up_8_p, a=1.2, v=0.25, r=0.05)
          $ 2341 "Spatula_otw" "breakAfter"
          movel(Spatula_otw_p, a=1.2, v=0.25)
          $ 2342 "switch_spat_S≔ False "
          global switch_spat_S=  False
        else:
          $ 2343 "ElseIf spatula≟'spatula_flat_M'"
          if (spatula == "spatula_flat_M"):
            $ 2344 "MoveJ"
            $ 2345 "Spatula_otw" "breakAfter"
            movej(get_inverse_kin(Spatula_otw_p, qnear=Spatula_otw_q), a=1.3962634015954636, v=1.0471975511965976)
            $ 2346 "spat_flatM_up" "breakAfter"
            movej(get_inverse_kin(spat_flatM_up_p, qnear=spat_flatM_up_q), a=1.3962634015954636, v=1.0471975511965976, r=0.05)
            $ 2347 "MoveL"
            $ 2348 "spat_flatM_pick" "breakAfter"
            movel(spat_flatM_pick_p, a=0.2, v=0.1)
            # begin: URCap Program Node
            #   Source: Robotiq_Grippers, 3.17.0.105337, Robotiq Inc.
            #   Type: Gripper
            $ 2349 "Gripper Open (1)"
            if not(gripper_connected[0]):
              popup("Gripper 1 must be connected to run this program.", "No connection", False, True, True)
            end
            if not(rq_is_gripper_activated("1")):
              popup("Gripper 1 is not activated. Go to Installation tab > Gripper to activate it and run the program again.", "Not activated", False, True, True)
            end
            rq_set_pos_spd_for(0, 128, 128, "1")
            rq_wait_pos_spe_for_request(0, 128, 128, "1")
            rq_go_to("1")
            rq_wait("1")
            # end: URCap Program Node
            $ 2350 "spat_flatM_up" "breakAfter"
            movel(spat_flatM_up_p, a=1.2, v=0.25, r=0.05)
            $ 2351 "Spatula_otw" "breakAfter"
            movel(Spatula_otw_p, a=1.2, v=0.25)
            $ 2352 "switch_spat_F_M≔ False "
            global switch_spat_F_M=  False
          else:
            $ 2353 "ElseIf spatula≟'spatula_flat_S'"
            if (spatula == "spatula_flat_S"):
              $ 2354 "MoveJ"
              $ 2355 "Spatula_otw" "breakAfter"
              movej(get_inverse_kin(Spatula_otw_p, qnear=Spatula_otw_q), a=1.3962634015954636, v=1.0471975511965976)
              $ 2356 "spat_flatS_up" "breakAfter"
              movej(get_inverse_kin(spat_flatS_up_p, qnear=spat_flatS_up_q), a=1.3962634015954636, v=1.0471975511965976, r=0.05)
              $ 2357 "MoveL"
              $ 2358 "spat_flatS_pick" "breakAfter"
              movel(spat_flatS_pick_p, a=0.2, v=0.1)
              # begin: URCap Program Node
              #   Source: Robotiq_Grippers, 3.17.0.105337, Robotiq Inc.
              #   Type: Gripper
              $ 2359 "Gripper Open (1)"
              if not(gripper_connected[0]):
                popup("Gripper 1 must be connected to run this program.", "No connection", False, True, True)
              end
              if not(rq_is_gripper_activated("1")):
                popup("Gripper 1 is not activated. Go to Installation tab > Gripper to activate it and run the program again.", "Not activated", False, True, True)
              end
              rq_set_pos_spd_for(0, 128, 128, "1")
              rq_wait_pos_spe_for_request(0, 128, 128, "1")
              rq_go_to("1")
              rq_wait("1")
              # end: URCap Program Node
              $ 2360 "spat_flatS_up" "breakAfter"
              movel(spat_flatS_up_p, a=1.2, v=0.25, r=0.05)
              $ 2361 "Spatula_otw" "breakAfter"
              movel(Spatula_otw_p, a=1.2, v=0.25)
              $ 2362 "switch_spat_F_S≔ False "
              global switch_spat_F_S=  False
            end
          end
        end
      end
    end
    $ 2363 "switch_spat_M≔ True "
    global switch_spat_M=  True
    $ 2364 "switch_spat_S≔ True "
    global switch_spat_S=  True
    $ 2365 "switch_spat_F_M≔ True "
    global switch_spat_F_M=  True
    $ 2366 "switch_spat_F_S≔ True "
    global switch_spat_F_S=  True
    $ 2367 "correction_reset()"
    correction_reset()
  elif (38 == switch_1):
    $ 2563 "Case 38"
    $ 2564 "Decap Powder container"
    $ 2565 "MoveJ"
    $ 2567 "Waypoint_7" "breakAfter"
    movej(get_inverse_kin(Waypoint_7_p, qnear=Waypoint_7_q), a=1.3962634015954636, v=1.0471975511965976, r=0.05)
    $ 2568 "MoveL"
    $ 2570 "Waypoint_8" "breakAfter"
    movel(Waypoint_8_p, a=1.2, v=0.25)
    $ 2571 "MoveL"
    $ 2572 "Decapp_above_3" "breakAfter"
    movel(Decapp_above_3_p, a=1.2, v=0.25)
    $ 2573 "Set GRP_3F_Open=On"
    set_standard_digital_out(5, True)
    $ 2574 "Wait: 0.5"
    sleep(0.5)
    $ 2575 "Decapp_place_3" "breakAfter"
    movel(Decapp_place_3_p, a=0.3, v=0.05)
    $ 2576 "Set GRP_3F_Open=Off"
    set_standard_digital_out(5, False)
    $ 2577 "Wait: 0.5"
    sleep(0.5)
    # begin: URCap Program Node
    #   Source: Robotiq_Grippers, 3.17.0.105337, Robotiq Inc.
    #   Type: Gripper
    $ 2578 "Gripper Open (1)"
    if not(gripper_connected[0]):
      popup("Gripper 1 must be connected to run this program.", "No connection", False, True, True)
    end
    if not(rq_is_gripper_activated("1")):
      popup("Gripper 1 is not activated. Go to Installation tab > Gripper to activate it and run the program again.", "Not activated", False, True, True)
    end
    rq_set_pos_spd_for(0, 77, 77, "1")
    rq_wait_pos_spe_for_request(0, 77, 77, "1")
    rq_go_to("1")
    rq_wait("1")
    # end: URCap Program Node
    $ 2579 "MoveL"
    $ 2580 "Decapp_above_4" "breakAfter"
    movel(Decapp_above_4_p, a=1.2, v=0.25)
    $ 2581 "Waypoint_78" "breakAfter"
    movel(Waypoint_78_p, a=1.2, v=0.25, r=0.05)
    $ 2582 "Home (Safe)"
    movej([-1.2302089344500047, -1.2969853503591224, -1.875639182904262, -1.539621866126728, 1.5731943360401213, -2.80099559440227], a=1.3962634015954636, v=1.0471975511965976)
  elif (39 == switch_1):
    $ 2583 "Case 39"
    $ 2584 "Powder container Pick"
    $ 2585 "Direct Pick"
    $ 2586 "Set"
    set_tcp(p[0.0,0.0,0.15052000000000001,3.1415,0.0,0.0])
    $ 2587 "read_db_data()"
    read_db_data()
    # begin: URCap Program Node
    #   Source: SensoPart VISOR Robotic, 2.0.6, SensoPart Industriesensorik GmbH
    #   Type: VISOR ChangeJob
    $ 2588 "# 1 VISOR ChangeJob"
    visor_changeJob(1, "Aztec_no_dot_pick", 6000)
    # end: URCap Program Node
    # begin: URCap Program Node
    #   Source: SensoPart VISOR Robotic, 2.0.6, SensoPart Industriesensorik GmbH
    #   Type: VISOR Terminal
    $ 2589 "# 1 VISOR Terminal"
    visor_terminal(1, "TRX00", 3000)
    # end: URCap Program Node
    $ 2590 "table_pick_TCP≔visor_getPose3d(1, 0)"
    global table_pick_TCP= visor_getPose3d (1, 0)
    # begin: URCap Program Node
    #   Source: Robotiq_Grippers, 3.17.0.105337, Robotiq Inc.
    #   Type: Gripper
    $ 2591 "Gripper Open (1)"
    if not(gripper_connected[0]):
      popup("Gripper 1 must be connected to run this program.", "No connection", False, True, True)
    end
    if not(rq_is_gripper_activated("1")):
      popup("Gripper 1 is not activated. Go to Installation tab > Gripper to activate it and run the program again.", "Not activated", False, True, True)
    end
    rq_set_pos_spd_for(0, 77, 77, "1")
    rq_wait_pos_spe_for_request(0, 77, 77, "1")
    rq_go_to("1")
    rq_wait("1")
    # end: URCap Program Node
    $ 2592 "MoveJ"
    $ 2594 "Waypoint_10" "breakAfter"
    movej(get_inverse_kin(Waypoint_10_p, qnear=Waypoint_10_q), a=1.3962634015954636, v=1.0471975511965976, r=0.05)
    $ 2595 "Waypoint_9" "breakAfter"
    movej(get_inverse_kin(Waypoint_9_p, qnear=Waypoint_9_q), a=1.3962634015954636, v=1.0471975511965976, r=0.05)
    $ 2596 "MoveJ"
    $ 2598 "table_prepick≔pose_trans(table_pick_TCP,p[0,0,cent_edge/2,0,0,0])"
    global table_prepick=pose_trans(table_pick_TCP,p[0,0,cent_edge/2,0,0,0])
    $ 2599 "table_prepick" "breakAfter"
    movej(table_prepick, a=0.8726646259971648, v=0.6981317007977318)
    $ 2600 "table_safe_pick≔pose_trans(table_prepick, p[0,pick_2_base-H_c,cent_edge/2,0,0,0])"
    global table_safe_pick= pose_trans (table_prepick, p[0,pick_2_base-H_c,cent_edge/2,0,0,0])
    $ 2601 "table_safe_pick" "breakAfter"
    movej(table_safe_pick, a=0.8726646259971648, v=0.6981317007977318, r=0.05)
    $ 2602 "table_pick≔pose_trans(table_prepick, p[0,pick_2_base - d_cc,0,0,0,0])"
    global table_pick= pose_trans (table_prepick, p[0,pick_2_base - d_cc,0,0,0,0])
    $ 2603 "table_pick" "breakAfter"
    movej(table_pick, a=0.8726646259971648, v=0.6981317007977318)
    # begin: URCap Program Node
    #   Source: Robotiq_Grippers, 3.17.0.105337, Robotiq Inc.
    #   Type: Gripper
    $ 2604 "Gripper Close (1)"
    if not(gripper_connected[0]):
      popup("Gripper 1 must be connected to run this program.", "No connection", False, True, True)
    end
    if not(rq_is_gripper_activated("1")):
      popup("Gripper 1 is not activated. Go to Installation tab > Gripper to activate it and run the program again.", "Not activated", False, True, True)
    end
    rq_set_pos_spd_for(255, 77, 51, "1")
    rq_wait_pos_spe_for_request(255, 77, 51, "1")
    rq_go_to("1")
    rq_wait("1")
    # end: URCap Program Node
    $ 2605 "table_prepick" "breakAfter"
    movej(table_prepick, a=0.8726646259971648, v=0.6981317007977318)
    $ 2606 "Picking≔ True "
    global Picking=  True
    $ 2608 "powder_position≔'Position2'"
    global powder_position="Position2"
    $ 2609 "MoveJ"
    $ 2610 "Powder_wayp1" "breakAfter"
    movej(get_inverse_kin(Powder_wayp1_p, qnear=Powder_wayp1_q), a=1.3962634015954636, v=1.0471975511965976, r=0.05)
    $ 2611 "MoveL"
    $ 2612 "Waypoint_2" "breakAfter"
    movel(Waypoint_2_p, a=1.2, v=0.25)
    $ 2613 "Set"
    set_tcp(p[0.0,0.0,0.161,3.1415,0.0,0.0])
    $ 2614 "If powder_position ≟ 'Position1'"
    if (powder_position  ==  "Position1"):
      $ 2615 "MoveJ"
      $ 2616 "Postions_otw" "breakAfter"
      movej(get_inverse_kin(Postions_otw_p, qnear=Postions_otw_q), a=1.3962634015954636, v=1.0471975511965976, r=0.01)
      $ 2617 "MoveL"
      $ 2618 "Cont_A_TCP" "breakAfter"
      movel(Cont_A_TCP, a=0.5, v=0.2)
      $ 2619 "cont_A_prepick≔pose_trans(Cont_A_TCP, p[0,0,cent_edge/2,0,0,0])"
      global cont_A_prepick= pose_trans (Cont_A_TCP, p[0,0,cent_edge/2,0,0,0])
      $ 2620 "cont_A_prepick" "breakAfter"
      movel(cont_A_prepick, a=0.3, v=0.05)
      $ 2621 "cont_A_pick≔pose_trans(cont_A_prepick, p[0,pick_2_base-d_cc,0,0,0,0])"
      global cont_A_pick= pose_trans (cont_A_prepick, p[0,pick_2_base-d_cc,0,0,0,0])
      $ 2622 "cont_A_pick" "breakAfter"
      movel(cont_A_pick, a=0.2, v=0.1)
      # begin: URCap Program Node
      #   Source: Robotiq_Grippers, 3.17.0.105337, Robotiq Inc.
      #   Type: Gripper
      $ 2623 "Gripper Open (1)"
      if not(gripper_connected[0]):
        popup("Gripper 1 must be connected to run this program.", "No connection", False, True, True)
      end
      if not(rq_is_gripper_activated("1")):
        popup("Gripper 1 is not activated. Go to Installation tab > Gripper to activate it and run the program again.", "Not activated", False, True, True)
      end
      rq_set_pos_spd_for(0, 77, 26, "1")
      rq_wait_pos_spe_for_request(0, 77, 26, "1")
      rq_go_to("1")
      rq_wait("1")
      # end: URCap Program Node
      $ 2624 "cont_A_otw" "breakAfter"
      movel(cont_A_otw_p, a=0.5, v=0.2)
      $ 2625 "cont_A_prepick" "breakAfter"
      movel(cont_A_prepick, a=0.5, v=0.2)
      $ 2626 "Postions_otw" "breakAfter"
      movel(Postions_otw_p, a=0.5, v=0.2, r=0.01)
      $ 2628 "Home (Safe)"
      movej([-1.2302089344500047, -1.2969853503591224, -1.875639182904262, -1.539621866126728, 1.5731943360401213, -2.80099559440227], a=1.3962634015954636, v=1.0471975511965976)
    else:
      $ 2630 "ElseIf powder_position≟'Position2'"
      if (powder_position == "Position2"):
        $ 2631 "MoveJ"
        $ 2632 "Postions_otw" "breakAfter"
        movej(get_inverse_kin(Postions_otw_p, qnear=Postions_otw_q), a=1.3962634015954636, v=1.0471975511965976, r=0.01)
        $ 2633 "MoveL"
        $ 2636 "cont_B_prepick≔pose_trans(Cont_B_TCP, p[0,0,cent_edge/2,0,0,0])"
        global cont_B_prepick= pose_trans (Cont_B_TCP, p[0,0,cent_edge/2,0,0,0])
        $ 2637 "cont_B_prepick" "breakAfter"
        movel(cont_B_prepick, a=1.2, v=0.25)
        $ 2638 "cont_B_pick≔pose_trans(cont_B_prepick, p[0,pick_2_base-d_cc,0,0,0,0])"
        global cont_B_pick= pose_trans (cont_B_prepick, p[0,pick_2_base-d_cc,0,0,0,0])
        $ 2639 "cont_B_pick" "breakAfter"
        global move_thread_flag_2639=0
        thread move_thread_2639():
          enter_critical
          move_thread_flag_2639 = 1
          movel(cont_B_pick, a=0.2, v=0.1)
          move_thread_flag_2639 = 2
          exit_critical
        end
        move_thread_flag_2639 = 0
        move_thread_han_2639 = run move_thread_2639()
        while (True):
          local targetTcpDirection=get_target_tcp_speed()
          local stepsToRetract=tool_contact(direction=targetTcpDirection, force_threshold=8.000000)
          if (stepsToRetract > 0):
            kill move_thread_han_2639
            stopl(3.0)
            local backTrackMovement=get_actual_joint_positions_history(stepsToRetract)
            local contactPose=get_forward_kin(backTrackMovement)
            local posDir=[targetTcpDirection[0],targetTcpDirection[1],targetTcpDirection[2]]
            local retractTo=contactPose
            if (norm(posDir) > 1e-6):
              local normalizedPosDir=normalize(posDir)
              local additionalRetraction=p[normalizedPosDir[0] * 0.0, normalizedPosDir[1] * 0.0, normalizedPosDir[2] * 0.0, 0, 0, 0]
              retractTo = pose_sub(contactPose, additionalRetraction)
            end
            movel(retractTo, a=3.0, v=0.1)
            $ 2640 "Until (tool_contact_detection)"
            $ 2641 "saved_place_pos≔get_actual_tcp_pose()"
            global saved_place_pos= get_actual_tcp_pose ()
            break
          end
          sleep(1.0E-10)
          if (move_thread_flag_2639 > 1):
            join move_thread_han_2639
            break
          end
          sync()
        end
        # begin: URCap Program Node
        #   Source: Robotiq_Grippers, 3.17.0.105337, Robotiq Inc.
        #   Type: Gripper
        $ 2642 "Gripper Open (1)"
        if not(gripper_connected[0]):
          popup("Gripper 1 must be connected to run this program.", "No connection", False, True, True)
        end
        if not(rq_is_gripper_activated("1")):
          popup("Gripper 1 is not activated. Go to Installation tab > Gripper to activate it and run the program again.", "Not activated", False, True, True)
        end
        rq_set_pos_spd_for(0, 77, 26, "1")
        rq_wait_pos_spe_for_request(0, 77, 26, "1")
        rq_go_to("1")
        rq_wait("1")
        # end: URCap Program Node
        $ 2643 "cont_B_otw" "breakAfter"
        movel(cont_B_otw_p, a=1.2, v=0.25)
        $ 2645 "cont_B_safe" "breakAfter"
        movel(cont_B_safe_p, a=1.2, v=0.25)
        $ 2646 "Postions_otw" "breakAfter"
        movel(Postions_otw_p, a=1.2, v=0.25)
        $ 2647 "Home (Safe)"
        movej([-1.2302089344500047, -1.2969853503591224, -1.875639182904262, -1.539621866126728, 1.5731943360401213, -2.80099559440227], a=1.3962634015954636, v=1.0471975511965976)
      else:
        $ 2649 "ElseIf powder_position≟'Position3'"
        if (powder_position == "Position3"):
          $ 2650 "MoveJ"
          $ 2651 "Postions_otw" "breakAfter"
          movej(get_inverse_kin(Postions_otw_p, qnear=Postions_otw_q), a=1.3962634015954636, v=1.0471975511965976, r=0.01)
          $ 2658 "MoveL"
          $ 2659 "Cont_C_TCP" "breakAfter"
          movel(Cont_C_TCP, a=1.2, v=0.25, r=0.01)
          $ 2660 "cont_C_prepick≔pose_trans(Cont_C_TCP, p[0,0,cent_edge/2,0,0,0])"
          global cont_C_prepick= pose_trans (Cont_C_TCP, p[0,0,cent_edge/2,0,0,0])
          $ 2661 "cont_C_prepick" "breakAfter"
          movel(cont_C_prepick, a=0.3, v=0.05)
          $ 2662 "cont_C_pick≔pose_trans(cont_C_prepick, p[0,pick_2_base-d_cc,0,0,0,0])"
          global cont_C_pick= pose_trans (cont_C_prepick, p[0,pick_2_base-d_cc,0,0,0,0])
          $ 2663 "cont_C_pick" "breakAfter"
          movel(cont_C_pick, a=0.2, v=0.1)
          # begin: URCap Program Node
          #   Source: Robotiq_Grippers, 3.17.0.105337, Robotiq Inc.
          #   Type: Gripper
          $ 2664 "Gripper Open (1)"
          if not(gripper_connected[0]):
            popup("Gripper 1 must be connected to run this program.", "No connection", False, True, True)
          end
          if not(rq_is_gripper_activated("1")):
            popup("Gripper 1 is not activated. Go to Installation tab > Gripper to activate it and run the program again.", "Not activated", False, True, True)
          end
          rq_set_pos_spd_for(0, 77, 26, "1")
          rq_wait_pos_spe_for_request(0, 77, 26, "1")
          rq_go_to("1")
          rq_wait("1")
          # end: URCap Program Node
          $ 2665 "cont_C_otw" "breakAfter"
          movel(cont_C_otw_p, a=1.2, v=0.25)
          $ 2666 "cont_C_prepick" "breakAfter"
          movel(cont_C_prepick, a=1.2, v=0.25, r=0.01)
          $ 2667 "Postions_otw" "breakAfter"
          movel(Postions_otw_p, a=1.2, v=0.25)
          $ 2668 "Home (Safe)"
          movej([-1.2302089344500047, -1.2969853503591224, -1.875639182904262, -1.539621866126728, 1.5731943360401213, -2.80099559440227], a=1.3962634015954636, v=1.0471975511965976)
        end
      end
    end
    $ 2670 "Home (Safe)"
    movej([-1.2302089344500047, -1.2969853503591224, -1.875639182904262, -1.539621866126728, 1.5731943360401213, -2.80099559440227], a=1.3962634015954636, v=1.0471975511965976)
  elif (41 == switch_1):
    $ 2779 "Case 41"
    $ 2780 "Task≔'Decapping_Dosing'"
    global Task="Decapping_Dosing"
    $ 2781 "tilt_to_home()"
    tilt_to_home()
    $ 2782 "Weigh, Place & decap container"
    $ 2783 "Set"
    set_tcp(p[0.0,0.0,0.15052000000000001,3.1415,0.0,0.0])
    # begin: URCap Program Node
    #   Source: SensoPart VISOR Robotic, 2.0.6, SensoPart Industriesensorik GmbH
    #   Type: VISOR Robotic App
    $ 2784 "VISOR Easy Pick"
    def visorFuncEasyPick_6a96fc():
      # begin: URCap Program Node
      #   Source: SensoPart VISOR Robotic, 2.0.6, SensoPart Industriesensorik GmbH
      #   Type: Easy Pick Setup
      $ 2785 "# 1 Setup" "noBreak"
      local easyPickVisorId = 1
      local easyPickArmMounted = True
      local easyPickSetJob = True
      local easyPickJobName = "PoTS"
      local easyPickAtImgAcq = False
      local easyPickImgAcqPose = FRM_PoTS
      # end: URCap Program Node
      # begin: URCap Program Node
      #   Source: SensoPart VISOR Robotic, 2.0.6, SensoPart Industriesensorik GmbH
      #   Type: Process
      $ 2786 "Process" "noBreak"
      local easyPickObjTaken = False
      local easyPickTrigger = False
      local easyPickPoseIdx = 0
      local easyPickPose = p[0,0,0,0,0,0]
      def easyPickFuncTrigger(visorId, setJob, jobName, arm):
      if (setJob):
        visor_changeJob(visorId, jobName, 6000)
      end
      if (arm):
        visor_trigger(visorId, 6000, "arm")
      else:
        visor_trigger(visorId, 6000)
      end
      global easyPickParts_7=visor_partsFound(visorId)
      visor_easyPickUpdate(visorId, "parts", visor_partsFound(visorId))
      return visor_getPose3d(visorId, 0)
    end
    while (not easyPickObjTaken):
      easyPickTrigger = (easyPickCount_7 >= visor_partsFound(easyPickVisorId)) or (easyPickCount_7 > 9) or (not visor_easyPickCheckIdent("eaa5b7", easyPickVisorId))
      if (easyPickTrigger):
        easyPickCount_7 = 0
      end
      easyPickPoseIdx = easyPickCount_7
      easyPickPose = visor_getPose3d(easyPickVisorId, easyPickPoseIdx)
      visor_easyPickUpdate(easyPickVisorId, "counter", easyPickPoseIdx)
      # begin: URCap Program Node
      #   Source: SensoPart VISOR Robotic, 2.0.6, SensoPart Industriesensorik GmbH
      #   Type: Image Acquisition Pose
      $ 2787 "Image Acquisition Pose" "noBreak"
      if (easyPickTrigger):
        if (not easyPickAtImgAcq):
          movej(pose_trans(easyPickImgAcqPose,p[0.0000,0.0000,-0.0000,0.0000,0.0000,0.0000]),a=1.3963,v=1.0472,t=0.000000,r=0.000000)
          easyPickAtImgAcq = True
        end
        easyPickPose = easyPickFuncTrigger(easyPickVisorId, easyPickSetJob, easyPickJobName, easyPickArmMounted)
      end
      # end: URCap Program Node
      # begin: URCap Program Node
      #   Source: SensoPart VISOR Robotic, 2.0.6, SensoPart Industriesensorik GmbH
      #   Type: Object Detected
      $ 2788 "Object Detected" "noBreak"
      if (visor_partsFound(easyPickVisorId) > 0):
        $ 2789 "Open Gripper" "noBreak"
        # begin: URCap Program Node
        #   Source: Robotiq_Grippers, 3.17.0.105337, Robotiq Inc.
        #   Type: Gripper
        $ 2790 "Gripper Open (1)" "noBreak"
        if not(gripper_connected[0]):
          popup("Gripper 1 must be connected to run this program.", "No connection", False, True, True)
        end
        if not(rq_is_gripper_activated("1")):
          popup("Gripper 1 is not activated. Go to Installation tab > Gripper to activate it and run the program again.", "Not activated", False, True, True)
        end
        rq_set_pos_spd_for(0, 77, 77, "1")
        rq_wait_pos_spe_for_request(0, 77, 77, "1")
        rq_go_to("1")
        rq_wait("1")
        # end: URCap Program Node
        $ 2791 "Set" "noBreak"
        set_tcp(p[0.0,0.0,0.161,3.1415,0.0,0.0])
        $ 2792 "Wait: 0.2" "noBreak"
        sleep(0.2)
        $ 2793 "Place on second weigh scale" "noBreak"
        $ 2794 "MoveJ" "noBreak"
        $ 2795 "Waypoint_1" "noBreak"
        movej(get_inverse_kin(Waypoint_1_p, qnear=Waypoint_1_q), a=1.3962634015954636, v=1.0471975511965976, r=0.1)
        $ 2796 "Waypoint_5" "noBreak"
        movej(get_inverse_kin(Waypoint_5_p, qnear=Waypoint_5_q), a=1.3962634015954636, v=1.0471975511965976)
        $ 2798 "If Picking≟ True " "noBreak"
        if (Picking ==   True  ):
          $ 2799 "Pick from saved pose" "noBreak"
          $ 2800 "MoveL" "noBreak"
          $ 2801 "cont_B_safe" "noBreak"
          movel(cont_B_safe_p, a=0.2, v=0.1)
          $ 2802 "saved_place_pos" "noBreak"
          movel(saved_place_pos, a=1.2, v=0.25)
          # begin: URCap Program Node
          #   Source: Robotiq_Grippers, 3.17.0.105337, Robotiq Inc.
          #   Type: Gripper
          $ 2803 "Gripper Close (1)" "noBreak"
          if not(gripper_connected[0]):
            popup("Gripper 1 must be connected to run this program.", "No connection", False, True, True)
          end
          if not(rq_is_gripper_activated("1")):
            popup("Gripper 1 is not activated. Go to Installation tab > Gripper to activate it and run the program again.", "Not activated", False, True, True)
          end
          rq_set_pos_spd_for(255, 77, 26, "1")
          rq_wait_pos_spe_for_request(255, 77, 26, "1")
          rq_go_to("1")
          rq_wait("1")
          # end: URCap Program Node
          $ 2804 "cont_B_safe" "noBreak"
          movel(cont_B_safe_p, a=1.2, v=0.25)
          $ 2805 "Postions_otw" "noBreak"
          movel(Postions_otw_p, a=1.2, v=0.25)
        else:
          $ 2808 "Else" "noBreak"
          $ 2809 "read_db_data()" "noBreak"
          read_db_data()
          $ 2810 "Pick from B" "noBreak"
          $ 2811 "MoveL" "noBreak"
          $ 2813 "cont_B_safe" "noBreak"
          movel(cont_B_safe_p, a=1.2, v=0.25)
          $ 2814 "cont_B_prepick≔pose_trans(Cont_B_TCP, p[0,0,cent_edge/2,0,0,0])" "noBreak"
          global cont_B_prepick= pose_trans (Cont_B_TCP, p[0,0,cent_edge/2,0,0,0])
          $ 2815 "cont_B_otw" "noBreak"
          movel(cont_B_otw_p, a=1.2, v=0.25)
          $ 2817 "cont_B_pick≔pose_trans(cont_B_prepick, p[0,pick_2_base-d_cc,0,0,0,0])" "noBreak"
          global cont_B_pick= pose_trans (cont_B_prepick, p[0,pick_2_base-d_cc,0,0,0,0])
          $ 2818 "cont_B_pick" "noBreak"
          movel(cont_B_pick, a=0.2, v=0.1)
          # begin: URCap Program Node
          #   Source: Robotiq_Grippers, 3.17.0.105337, Robotiq Inc.
          #   Type: Gripper
          $ 2819 "Gripper Close (1)" "noBreak"
          if not(gripper_connected[0]):
            popup("Gripper 1 must be connected to run this program.", "No connection", False, True, True)
          end
          if not(rq_is_gripper_activated("1")):
            popup("Gripper 1 is not activated. Go to Installation tab > Gripper to activate it and run the program again.", "Not activated", False, True, True)
          end
          rq_set_pos_spd_for(255, 77, 51, "1")
          rq_wait_pos_spe_for_request(255, 77, 51, "1")
          rq_go_to("1")
          rq_wait("1")
          # end: URCap Program Node
          $ 2820 "cont_B_prepick" "noBreak"
          movel(cont_B_prepick, a=1.2, v=0.25, r=0.01)
          $ 2821 "Postions_otw" "noBreak"
          movel(Postions_otw_p, a=1.2, v=0.25)
        end
        $ 2838 "Set" "noBreak"
        set_tcp(p[0.0,0.0,0.15052000000000001,3.1415,0.0,0.0])
        # begin: URCap Program Node
        #   Source: SensoPart VISOR Robotic, 2.0.6, SensoPart Industriesensorik GmbH
        #   Type: Approach Pose
        $ 2839 "Approach Pose" "noBreak"
        movej(pose_trans(easyPickPose,p[0.0000,0.0000,-0.0000,0.0000,0.0000,0.0000]),a=0.5236,v=0.4363,t=0.000000,r=0.000000)
        # end: URCap Program Node
        # begin: URCap Program Node
        #   Source: SensoPart VISOR Robotic, 2.0.6, SensoPart Industriesensorik GmbH
        #   Type: Target Pose
        $ 2840 "Target Pose" "noBreak"
        movel(pose_trans(easyPickPose,p[0.0000,0.0000,-0.0000,0.0000,0.0000,0.0000]),a=0.1000,v=0.0500,t=0.000000,r=0.000000)
        # end: URCap Program Node
        $ 2841 "Close Gripper" "noBreak"
        $ 2842 "container_place≔get_actual_tcp_pose()" "noBreak"
        global container_place= get_actual_tcp_pose ()
        $ 2843 "PoTS_place_abov≔pose_trans(container_place, p[0,0,cent_edge/2,0,0,0])" "noBreak"
        global PoTS_place_abov=pose_trans(container_place, p[0,0,cent_edge/2,0,0,0])
        $ 2844 "MoveL" "noBreak"
        $ 2845 "PoTS_place_abov" "noBreak"
        movel(PoTS_place_abov, a=0.5, v=0.05)
        $ 2847 "target_pose≔pose_trans(PoTS_place_abov, p[0,pick_2_base-d_cc,0,0,0,0])" "noBreak"
        global target_pose=pose_trans(PoTS_place_abov, p[0,pick_2_base-d_cc,0,0,0,0])
        $ 2848 "MoveL" "noBreak"
        $ 2849 "target_pose" "noBreak"
        movel(target_pose, a=0.3, v=0.05)
        # begin: URCap Program Node
        #   Source: Robotiq_Grippers, 3.17.0.105337, Robotiq Inc.
        #   Type: Gripper
        $ 2850 "Gripper Open (1)" "noBreak"
        if not(gripper_connected[0]):
          popup("Gripper 1 must be connected to run this program.", "No connection", False, True, True)
        end
        if not(rq_is_gripper_activated("1")):
          popup("Gripper 1 is not activated. Go to Installation tab > Gripper to activate it and run the program again.", "Not activated", False, True, True)
        end
        rq_set_pos_spd_for(0, 77, 77, "1")
        rq_wait_pos_spe_for_request(0, 77, 77, "1")
        rq_go_to("1")
        rq_wait("1")
        # end: URCap Program Node
        # begin: URCap Program Node
        #   Source: SensoPart VISOR Robotic, 2.0.6, SensoPart Industriesensorik GmbH
        #   Type: Exit Pose
        $ 2851 "Exit Pose" "noBreak"
        movel(pose_trans(easyPickPose,p[0.0000,0.0000,0.1000,0.0000,0.0000,0.0000]),a=0.5000,v=0.2500,t=0.000000,r=0.000000)
        # end: URCap Program Node
        easyPickObjTaken = True
      end
      # end: URCap Program Node
      # begin: URCap Program Node
      #   Source: SensoPart VISOR Robotic, 2.0.6, SensoPart Industriesensorik GmbH
      #   Type: No Object Detected
      $ 2852 "No Object Detected" "noBreak"
      if (visor_partsFound(easyPickVisorId) < 1):
        $ 2853 "Popup: No POTS detected" "noBreak"
        popup("No POTS detected", "Message", False, False, blocking=True)
        else:
      end
      # end: URCap Program Node
    end
    easyPickCount_7 = easyPickCount_7 + 1
    visor_easyPickUpdate(easyPickVisorId, "counter", easyPickCount_7)
    visor_easyPickSetIdent("eaa5b7", easyPickVisorId)
    # end: URCap Program Node
  end
  visorFuncEasyPick_6a96fc()
  # end: URCap Program Node
  $ 2888 "MoveJ"
  $ 2889 "place_2_home" "breakAfter"
  movej(get_inverse_kin(place_2_home_p, qnear=place_2_home_q), a=1.3962634015954636, v=1.0471975511965976)
  $ 2890 "Picking≔ False "
  global Picking=  False
  elif (42 == switch_1):
    $ 2891 "Case 42"
  elif (43 == switch_1):
    $ 3653 "Case 43"
  elif (44 == switch_1):
    $ 3906 "Case 44"
  elif (45 == switch_1):
    $ 3970 "Case 45"
  elif (46 == switch_1):
    $ 4007 "Case 46"
  elif (47 == switch_1):
    $ 4297 "Case 47"
  elif (48 == switch_1):
    $ 4352 "Case 48"
  elif (49 == switch_1):
    $ 4370 "Case 49"
  elif (50 == switch_1):
    $ 4388 "Case 50"
    $ 4389 "Emptying powder container"
    $ 4390 "tilt_to_home()"
    tilt_to_home()
    $ 4391 "scoop_status≔'emptying'"
    global scoop_status="emptying"
    $ 4392 "Dosing untill empty"
    $ 4393 "tilt_angle_sent≔0.0"
    global tilt_angle_sent=0.0
    $ 4394 "send_target_info()"
    send_target_info()
    $ 4395 "zero_scale()"
    zero_scale()
    $ 4396 "prev_spat≔''"
    global prev_spat=""
    $ 4397 "spatula≔''"
    global spatula=""
    $ 4398 "send_powder_info()"
    send_powder_info()
    $ 4399 "Set AO[0]=0.0"
    set_standard_analog_out(0, 0.0)
    $ 4400 "Wait: 0.2"
    sleep(0.2)
    $ 4401 "reach pots decapping pose"
    # begin: URCap Program Node
    #   Source: SensoPart VISOR Robotic, 2.0.6, SensoPart Industriesensorik GmbH
    #   Type: VISOR Robotic App
    $ 4407 "VISOR Easy Pick"
    def visorFuncEasyPick_f946db():
      # begin: URCap Program Node
      #   Source: SensoPart VISOR Robotic, 2.0.6, SensoPart Industriesensorik GmbH
      #   Type: Easy Pick Setup
      $ 4408 "# 1 Setup" "noBreak"
      local easyPickVisorId = 1
      local easyPickArmMounted = True
      local easyPickSetJob = True
      local easyPickJobName = "Weight_scale"
      local easyPickAtImgAcq = False
      local easyPickImgAcqPose = Trigger
      # end: URCap Program Node
      # begin: URCap Program Node
      #   Source: SensoPart VISOR Robotic, 2.0.6, SensoPart Industriesensorik GmbH
      #   Type: Process
      $ 4409 "Process" "noBreak"
      local easyPickObjTaken = False
      local easyPickTrigger = False
      local easyPickPoseIdx = 0
      local easyPickPose = p[0,0,0,0,0,0]
      def easyPickFuncTrigger(visorId, setJob, jobName, arm):
      if (setJob):
        visor_changeJob(visorId, jobName, 6000)
      end
      if (arm):
        visor_trigger(visorId, 6000, "arm")
      else:
        visor_trigger(visorId, 6000)
      end
      global easyPickParts_4=visor_partsFound(visorId)
      visor_easyPickUpdate(visorId, "parts", visor_partsFound(visorId))
      return visor_getPose3d(visorId, 0)
    end
    while (not easyPickObjTaken):
      easyPickTrigger = (easyPickCount_4 >= visor_partsFound(easyPickVisorId)) or (easyPickCount_4 > 9) or (not visor_easyPickCheckIdent("be50ea", easyPickVisorId))
      if (easyPickTrigger):
        easyPickCount_4 = 0
      end
      easyPickPoseIdx = easyPickCount_4
      easyPickPose = visor_getPose3d(easyPickVisorId, easyPickPoseIdx)
      visor_easyPickUpdate(easyPickVisorId, "counter", easyPickPoseIdx)
      # begin: URCap Program Node
      #   Source: SensoPart VISOR Robotic, 2.0.6, SensoPart Industriesensorik GmbH
      #   Type: Image Acquisition Pose
      $ 4410 "Image Acquisition Pose" "noBreak"
      if (easyPickTrigger):
        if (not easyPickAtImgAcq):
          movej(pose_trans(easyPickImgAcqPose,p[0.0000,0.0000,-0.0000,0.0000,0.0000,0.0000]),a=1.3963,v=1.0472,t=0.000000,r=0.000000)
          easyPickAtImgAcq = True
        end
        easyPickPose = easyPickFuncTrigger(easyPickVisorId, easyPickSetJob, easyPickJobName, easyPickArmMounted)
      end
      # end: URCap Program Node
      # begin: URCap Program Node
      #   Source: SensoPart VISOR Robotic, 2.0.6, SensoPart Industriesensorik GmbH
      #   Type: Object Detected
      $ 4411 "Object Detected" "noBreak"
      if (visor_partsFound(easyPickVisorId) > 0):
        $ 4412 "Open Gripper" "noBreak"
        $ 4413 "weight_value≔get_weight()" "noBreak"
        global weight_value=get_weight()
        $ 4414 "Wait: 1.0" "noBreak"
        sleep(1.0)
        $ 4415 "diff≔target_weight-weight_value" "noBreak"
        global diff=target_weight-weight_value
        $ 4416 "compute_level_percent(W_now, weight_value)" "noBreak"
        compute_level_percent(W_now, weight_value)
        $ 4417 "send_level_info()" "noBreak"
        send_level_info()
        $ 4418 "spatula≔select_spatula(Flowability, level, diff, bulk_density, mouth_d)" "noBreak"
        global spatula=select_spatula(Flowability, level, diff, bulk_density, mouth_d)
        $ 4419 "Wait: 0.2" "noBreak"
        sleep(0.2)
        $ 4420 "send_spatula_info()" "noBreak"
        send_spatula_info()
        $ 4421 "Pick spatula" "noBreak"
        $ 4422 "If spatula ≟ 'spatula_L'" "noBreak"
        if (spatula  ==  "spatula_L"):
          $ 4423 "MoveJ" "noBreak"
          $ 4424 "Spatula_otw" "noBreak"
          movej(get_inverse_kin(Spatula_otw_p, qnear=Spatula_otw_q), a=1.3962634015954636, v=1.0471975511965976)
          $ 4425 "pick_spat_L_abv" "noBreak"
          movej(get_inverse_kin(pick_spat_L_abv_p, qnear=pick_spat_L_abv_q), a=1.3962634015954636, v=1.0471975511965976)
          $ 4426 "MoveL" "noBreak"
          $ 4427 "spat_L_pick" "noBreak"
          movel(spat_L_pick_p, a=1.2, v=0.25)
          # begin: URCap Program Node
          #   Source: Robotiq_Grippers, 3.17.0.105337, Robotiq Inc.
          #   Type: Gripper
          $ 4428 "Gripper Close (1)" "noBreak"
          if not(gripper_connected[0]):
            popup("Gripper 1 must be connected to run this program.", "No connection", False, True, True)
          end
          if not(rq_is_gripper_activated("1")):
            popup("Gripper 1 is not activated. Go to Installation tab > Gripper to activate it and run the program again.", "Not activated", False, True, True)
          end
          rq_set_pos_spd_for(255, 0, 77, "1")
          rq_wait_pos_spe_for_request(255, 0, 77, "1")
          rq_go_to("1")
          rq_wait("1")
          # end: URCap Program Node
          $ 4429 "spat_L_lift" "noBreak"
          movel(spat_L_lift_p, a=1.2, v=0.25, r=0.01)
          $ 4430 "spat_L_side" "noBreak"
          movel(spat_L_side_p, a=1.2, v=0.25, r=0.01)
          $ 4431 "spat_L_up" "noBreak"
          movel(spat_L_up_p, a=1.2, v=0.25, r=0.05)
          $ 4432 "MoveJ" "noBreak"
          $ 4433 "Spatula_otw" "noBreak"
          movej(get_inverse_kin(Spatula_otw_p, qnear=Spatula_otw_q), a=1.3962634015954636, v=1.0471975511965976)
        else:
          $ 4434 "ElseIf spatula ≟'spatula_M'" "noBreak"
          if (spatula  == "spatula_M"):
            $ 4435 "MoveJ" "noBreak"
            $ 4436 "Spatula_otw" "noBreak"
            movej(get_inverse_kin(Spatula_otw_p, qnear=Spatula_otw_q), a=1.3962634015954636, v=1.0471975511965976)
            $ 4437 "spat_M_up" "noBreak"
            movej(get_inverse_kin(spat_M_up_p, qnear=spat_M_up_q), a=1.3962634015954636, v=1.0471975511965976, r=0.05)
            $ 4438 "MoveL" "noBreak"
            $ 4439 "spat_M_pick" "noBreak"
            movel(spat_M_pick_p, a=1.2, v=0.25)
            # begin: URCap Program Node
            #   Source: Robotiq_Grippers, 3.17.0.105337, Robotiq Inc.
            #   Type: Gripper
            $ 4440 "Gripper Close (1)" "noBreak"
            if not(gripper_connected[0]):
              popup("Gripper 1 must be connected to run this program.", "No connection", False, True, True)
            end
            if not(rq_is_gripper_activated("1")):
              popup("Gripper 1 is not activated. Go to Installation tab > Gripper to activate it and run the program again.", "Not activated", False, True, True)
            end
            rq_set_pos_spd_for(255, 0, 77, "1")
            rq_wait_pos_spe_for_request(255, 0, 77, "1")
            rq_go_to("1")
            rq_wait("1")
            # end: URCap Program Node
            $ 4441 "spat_M_up" "noBreak"
            movel(spat_M_up_p, a=1.2, v=0.25, r=0.05)
            $ 4442 "Spatula_otw" "noBreak"
            movel(Spatula_otw_p, a=1.2, v=0.25)
            $ 4443 "switch_spat_M≔ False " "noBreak"
            global switch_spat_M=  False
          else:
            $ 4444 "ElseIf spatula≟'spatula_S'" "noBreak"
            if (spatula == "spatula_S"):
              $ 4445 "MoveJ" "noBreak"
              $ 4446 "Spatula_otw" "noBreak"
              movej(get_inverse_kin(Spatula_otw_p, qnear=Spatula_otw_q), a=1.3962634015954636, v=1.0471975511965976)
              $ 4447 "spat_S_Up_7" "noBreak"
              movej(get_inverse_kin(spat_S_Up_7_p, qnear=spat_S_Up_7_q), a=1.3962634015954636, v=1.0471975511965976, r=0.05)
              $ 4448 "MoveL" "noBreak"
              $ 4449 "spat_S_Pick_4" "noBreak"
              movel(spat_S_Pick_4_p, a=1.2, v=0.25)
              # begin: URCap Program Node
              #   Source: Robotiq_Grippers, 3.17.0.105337, Robotiq Inc.
              #   Type: Gripper
              $ 4450 "Gripper Close (1)" "noBreak"
              if not(gripper_connected[0]):
                popup("Gripper 1 must be connected to run this program.", "No connection", False, True, True)
              end
              if not(rq_is_gripper_activated("1")):
                popup("Gripper 1 is not activated. Go to Installation tab > Gripper to activate it and run the program again.", "Not activated", False, True, True)
              end
              rq_set_pos_spd_for(255, 0, 77, "1")
              rq_wait_pos_spe_for_request(255, 0, 77, "1")
              rq_go_to("1")
              rq_wait("1")
              # end: URCap Program Node
              $ 4451 "spat_S_Up_8" "noBreak"
              movel(spat_S_Up_8_p, a=1.2, v=0.25, r=0.05)
              $ 4452 "Spatula_otw" "noBreak"
              movel(Spatula_otw_p, a=1.2, v=0.25)
              $ 4453 "switch_spat_S≔ False " "noBreak"
              global switch_spat_S=  False
            else:
              $ 4454 "ElseIf spatula≟'spatula_flat_M'" "noBreak"
              if (spatula == "spatula_flat_M"):
                $ 4455 "MoveJ" "noBreak"
                $ 4456 "Spatula_otw" "noBreak"
                movej(get_inverse_kin(Spatula_otw_p, qnear=Spatula_otw_q), a=1.3962634015954636, v=1.0471975511965976)
                $ 4457 "spat_flatM_up" "noBreak"
                movej(get_inverse_kin(spat_flatM_up_p, qnear=spat_flatM_up_q), a=1.3962634015954636, v=1.0471975511965976, r=0.05)
                $ 4458 "MoveL" "noBreak"
                $ 4459 "spat_flatM_pick" "noBreak"
                movel(spat_flatM_pick_p, a=1.2, v=0.25)
                # begin: URCap Program Node
                #   Source: Robotiq_Grippers, 3.17.0.105337, Robotiq Inc.
                #   Type: Gripper
                $ 4460 "Gripper Close (1)" "noBreak"
                if not(gripper_connected[0]):
                  popup("Gripper 1 must be connected to run this program.", "No connection", False, True, True)
                end
                if not(rq_is_gripper_activated("1")):
                  popup("Gripper 1 is not activated. Go to Installation tab > Gripper to activate it and run the program again.", "Not activated", False, True, True)
                end
                rq_set_pos_spd_for(255, 0, 77, "1")
                rq_wait_pos_spe_for_request(255, 0, 77, "1")
                rq_go_to("1")
                rq_wait("1")
                # end: URCap Program Node
                $ 4461 "spat_flatM_up" "noBreak"
                movel(spat_flatM_up_p, a=1.2, v=0.25, r=0.05)
                $ 4462 "Spatula_otw" "noBreak"
                movel(Spatula_otw_p, a=1.2, v=0.25)
                $ 4463 "switch_spat_F_M≔ False " "noBreak"
                global switch_spat_F_M=  False
              else:
                $ 4464 "ElseIf spatula≟'spatula_flat_S'" "noBreak"
                if (spatula == "spatula_flat_S"):
                  $ 4465 "MoveJ" "noBreak"
                  $ 4466 "Spatula_otw" "noBreak"
                  movej(get_inverse_kin(Spatula_otw_p, qnear=Spatula_otw_q), a=1.3962634015954636, v=1.0471975511965976)
                  $ 4467 "spat_flatS_up" "noBreak"
                  movej(get_inverse_kin(spat_flatS_up_p, qnear=spat_flatS_up_q), a=1.3962634015954636, v=1.0471975511965976, r=0.05)
                  $ 4468 "MoveL" "noBreak"
                  $ 4469 "spat_flatS_pick" "noBreak"
                  movel(spat_flatS_pick_p, a=1.2, v=0.25)
                  # begin: URCap Program Node
                  #   Source: Robotiq_Grippers, 3.17.0.105337, Robotiq Inc.
                  #   Type: Gripper
                  $ 4470 "Gripper Close (1)" "noBreak"
                  if not(gripper_connected[0]):
                    popup("Gripper 1 must be connected to run this program.", "No connection", False, True, True)
                  end
                  if not(rq_is_gripper_activated("1")):
                    popup("Gripper 1 is not activated. Go to Installation tab > Gripper to activate it and run the program again.", "Not activated", False, True, True)
                  end
                  rq_set_pos_spd_for(255, 0, 77, "1")
                  rq_wait_pos_spe_for_request(255, 0, 77, "1")
                  rq_go_to("1")
                  rq_wait("1")
                  # end: URCap Program Node
                  $ 4471 "spat_flatS_up" "noBreak"
                  movel(spat_flatS_up_p, a=1.2, v=0.25, r=0.05)
                  $ 4472 "Spatula_otw" "noBreak"
                  movel(Spatula_otw_p, a=1.2, v=0.25)
                  $ 4473 "switch_spat_F_S≔ False " "noBreak"
                  global switch_spat_F_S=  False
                end
              end
            end
          end
        end
        $ 4474 "Action_Info≔'Scooping'" "noBreak"
        global Action_Info="Scooping"
        $ 4475 "auto_tilt_and_scoop(W_now, target_weight, weight_value)" "noBreak"
        auto_tilt_and_scoop(W_now, target_weight, weight_value)
        $ 4476 "Action_Info≔'Dosing'" "noBreak"
        global Action_Info="Dosing"
        # begin: URCap Program Node
        #   Source: SensoPart VISOR Robotic, 2.0.6, SensoPart Industriesensorik GmbH
        #   Type: Approach Pose
        $ 4477 "Approach Pose" "noBreak"
        movej(pose_trans(easyPickPose,p[0.0000,0.0000,-0.0000,0.0000,0.0000,0.0000]),a=0.2618,v=0.1745,t=0.000000,r=0.000000)
        # end: URCap Program Node
        # begin: URCap Program Node
        #   Source: SensoPart VISOR Robotic, 2.0.6, SensoPart Industriesensorik GmbH
        #   Type: Target Pose
        $ 4478 "Target Pose" "noBreak"
        movel(pose_trans(easyPickPose,p[0.0000,0.0000,-0.0000,0.0000,0.0000,0.0000]),a=0.0500,v=0.0200,t=0.000000,r=0.000000)
        # end: URCap Program Node
        $ 4479 "Close Gripper" "noBreak"
        $ 4480 "dispense_pos≔get_actual_tcp_pose()" "noBreak"
        global dispense_pos= get_actual_tcp_pose ()
        $ 4481 "Loop weight_value≤target_weight and delta_count<3" "noBreak"
        thread Thread_while_4481():
          while (True):
            $ 4482 "MoveL" "noBreak"
            $ 4483 "dispense_pos" "noBreak"
            movel(dispense_pos, a=0.2, v=0.1)
            $ 4484 "log_weight()" "noBreak"
            log_weight()
            $ 4485 "CCW_full_Rotate()" "noBreak"
            CCW_full_Rotate()
            $ 4486 "Wait: 0.5" "noBreak"
            sleep(0.5)
            $ 4487 "tilt_pose≔pose_trans(get_actual_tcp_pose(), p[0, 0, 0, 0, 0, 2.0])" "noBreak"
            global tilt_pose=pose_trans(get_actual_tcp_pose(), p[0, 0, 0, 0, 0, 2.0])
            $ 4488 "movel(tilt_pose, a=0.5, v=0.5, r=0.00001)" "noBreak"
            movel(tilt_pose, a=0.5, v=0.5, r=0.00001)
            $ 4489 "weight_value≔get_weight()" "noBreak"
            global weight_value=get_weight()
            $ 4490 "tilt_angle≔-1" "noBreak"
            global tilt_angle=-1
            $ 4491 "Wait: 0.5" "noBreak"
            sleep(0.5)
            $ 4492 "dispense_pos" "noBreak"
            movel(dispense_pos, a=1.2, v=0.25)
            $ 4493 "compute_level_percent(W_now, weight_value)" "noBreak"
            compute_level_percent(W_now, weight_value)
            $ 4494 "If delta<0.01" "noBreak"
            if (delta<0.01):
              $ 4495 "delta_count≔delta_count+1" "noBreak"
              global delta_count=delta_count+1
            else:
              $ 4496 "Else" "noBreak"
              $ 4497 "delta_count≔0" "noBreak"
              global delta_count=0
            end
            $ 4498 "prev_spat≔spatula" "noBreak"
            global prev_spat=spatula
            $ 4499 "Wait: 0.2" "noBreak"
            sleep(0.2)
            $ 4500 "spatula≔select_spatula(Flowability, level, diff, bulk_density, mouth_d)" "noBreak"
            global spatula=select_spatula(Flowability, level, diff, bulk_density, mouth_d)
            $ 4501 "Wait: 1.0" "noBreak"
            sleep(1.0)
            $ 4502 "send_level_info()" "noBreak"
            send_level_info()
            $ 4503 "send_spatula_info()" "noBreak"
            send_spatula_info()
            $ 4504 "Set AO[0]=0.0" "noBreak"
            set_standard_analog_out(0, 0.0)
            $ 4505 "Wait: 0.5" "noBreak"
            sleep(0.5)
            $ 4506 "swtich spatula" "noBreak"
            $ 4507 "If spatula ≟ 'spatula_M' and switch_spat_M≟ True " "noBreak"
            if (spatula  ==  "spatula_M"  and  switch_spat_M ==   True  ):
              $ 4508 "MoveJ" "noBreak"
              $ 4509 "Spatula_otw" "noBreak"
              movej(get_inverse_kin(Spatula_otw_p, qnear=Spatula_otw_q), a=1.3962634015954636, v=1.0471975511965976)
              $ 4510 "spat_L_up" "noBreak"
              movej(get_inverse_kin(spat_L_up_p, qnear=spat_L_up_q), a=1.3962634015954636, v=1.0471975511965976)
              $ 4511 "MoveL" "noBreak"
              $ 4512 "spat_L_side" "noBreak"
              movel(spat_L_side_p, a=1.2, v=0.25)
              $ 4513 "spat_L_lift" "noBreak"
              movel(spat_L_lift_p, a=1.2, v=0.25)
              $ 4514 "spat_L_pick" "noBreak"
              movel(spat_L_pick_p, a=0.2, v=0.1)
              # begin: URCap Program Node
              #   Source: Robotiq_Grippers, 3.17.0.105337, Robotiq Inc.
              #   Type: Gripper
              $ 4515 "Gripper Open (1)" "noBreak"
              if not(gripper_connected[0]):
                popup("Gripper 1 must be connected to run this program.", "No connection", False, True, True)
              end
              if not(rq_is_gripper_activated("1")):
                popup("Gripper 1 is not activated. Go to Installation tab > Gripper to activate it and run the program again.", "Not activated", False, True, True)
              end
              rq_set_pos_spd_for(0, 255, 77, "1")
              rq_wait_pos_spe_for_request(0, 255, 77, "1")
              rq_go_to("1")
              rq_wait("1")
              # end: URCap Program Node
              $ 4516 "spat_M_pick" "noBreak"
              movel(spat_M_pick_p, a=1.2, v=0.25)
              # begin: URCap Program Node
              #   Source: Robotiq_Grippers, 3.17.0.105337, Robotiq Inc.
              #   Type: Gripper
              $ 4517 "Gripper Close (1)" "noBreak"
              if not(gripper_connected[0]):
                popup("Gripper 1 must be connected to run this program.", "No connection", False, True, True)
              end
              if not(rq_is_gripper_activated("1")):
                popup("Gripper 1 is not activated. Go to Installation tab > Gripper to activate it and run the program again.", "Not activated", False, True, True)
              end
              rq_set_pos_spd_for(255, 0, 77, "1")
              rq_wait_pos_spe_for_request(255, 0, 77, "1")
              rq_go_to("1")
              rq_wait("1")
              # end: URCap Program Node
              $ 4518 "spat_M_up" "noBreak"
              movel(spat_M_up_p, a=1.2, v=0.25)
              $ 4519 "Spatula_otw" "noBreak"
              movel(Spatula_otw_p, a=1.2, v=0.25)
              $ 4520 "switch_spat_M≔ False " "noBreak"
              global switch_spat_M=  False
              $ 4521 "correction_reset()" "noBreak"
              correction_reset()
            else:
              $ 4522 "ElseIf spatula ≟ 'spatula_S' and switch_spat_S ≟ True and prev_spat≟'spatula_M'" "noBreak"
              if (spatula  ==  "spatula_S" and switch_spat_S  ==   True  and prev_spat == "spatula_M"):
                $ 4523 "MoveL" "noBreak"
                $ 4524 "Spatula_otw" "noBreak"
                movel(Spatula_otw_p, a=1.2, v=0.25)
                $ 4525 "spat_M_up" "noBreak"
                movel(spat_M_up_p, a=1.2, v=0.25)
                $ 4526 "spat_M_pick" "noBreak"
                movel(spat_M_pick_p, a=0.2, v=0.1)
                # begin: URCap Program Node
                #   Source: Robotiq_Grippers, 3.17.0.105337, Robotiq Inc.
                #   Type: Gripper
                $ 4527 "Gripper Open (1)" "noBreak"
                if not(gripper_connected[0]):
                  popup("Gripper 1 must be connected to run this program.", "No connection", False, True, True)
                end
                if not(rq_is_gripper_activated("1")):
                  popup("Gripper 1 is not activated. Go to Installation tab > Gripper to activate it and run the program again.", "Not activated", False, True, True)
                end
                rq_set_pos_spd_for(0, 255, 77, "1")
                rq_wait_pos_spe_for_request(0, 255, 77, "1")
                rq_go_to("1")
                rq_wait("1")
                # end: URCap Program Node
                $ 4528 "spat_S_pick" "noBreak"
                movel(spat_S_pick_p, a=1.2, v=0.25)
                # begin: URCap Program Node
                #   Source: Robotiq_Grippers, 3.17.0.105337, Robotiq Inc.
                #   Type: Gripper
                $ 4529 "Gripper Close (1)" "noBreak"
                if not(gripper_connected[0]):
                  popup("Gripper 1 must be connected to run this program.", "No connection", False, True, True)
                end
                if not(rq_is_gripper_activated("1")):
                  popup("Gripper 1 is not activated. Go to Installation tab > Gripper to activate it and run the program again.", "Not activated", False, True, True)
                end
                rq_set_pos_spd_for(255, 0, 77, "1")
                rq_wait_pos_spe_for_request(255, 0, 77, "1")
                rq_go_to("1")
                rq_wait("1")
                # end: URCap Program Node
                $ 4530 "spat_S_up" "noBreak"
                movel(spat_S_up_p, a=1.2, v=0.25)
                $ 4531 "Spatula_otw" "noBreak"
                movel(Spatula_otw_p, a=1.2, v=0.25)
                $ 4532 "switch_spat_S≔ False " "noBreak"
                global switch_spat_S=  False
                $ 4533 "correction_reset()" "noBreak"
                correction_reset()
              else:
                $ 4534 "ElseIf spatula≟'spatula_S' and switch_spat_S≟ True  and prev_spat≟'spatula_L'" "noBreak"
                if (spatula == "spatula_S" and switch_spat_S ==   True    and  prev_spat == "spatula_L"):
                  $ 4535 "MoveJ" "noBreak"
                  $ 4536 "Spatula_otw" "noBreak"
                  movej(get_inverse_kin(Spatula_otw_p, qnear=Spatula_otw_q), a=1.3962634015954636, v=1.0471975511965976)
                  $ 4537 "spat_L_up" "noBreak"
                  movej(get_inverse_kin(spat_L_up_p, qnear=spat_L_up_q), a=1.3962634015954636, v=1.0471975511965976)
                  $ 4538 "MoveL" "noBreak"
                  $ 4539 "spat_L_side" "noBreak"
                  movel(spat_L_side_p, a=1.2, v=0.25)
                  $ 4540 "spat_L_lift" "noBreak"
                  movel(spat_L_lift_p, a=1.2, v=0.25)
                  $ 4541 "spat_L_pick" "noBreak"
                  movel(spat_L_pick_p, a=0.2, v=0.1)
                  # begin: URCap Program Node
                  #   Source: Robotiq_Grippers, 3.17.0.105337, Robotiq Inc.
                  #   Type: Gripper
                  $ 4542 "Gripper Open (1)" "noBreak"
                  if not(gripper_connected[0]):
                    popup("Gripper 1 must be connected to run this program.", "No connection", False, True, True)
                  end
                  if not(rq_is_gripper_activated("1")):
                    popup("Gripper 1 is not activated. Go to Installation tab > Gripper to activate it and run the program again.", "Not activated", False, True, True)
                  end
                  rq_set_pos_spd_for(0, 255, 77, "1")
                  rq_wait_pos_spe_for_request(0, 255, 77, "1")
                  rq_go_to("1")
                  rq_wait("1")
                  # end: URCap Program Node
                  $ 4543 "spat_S_pick" "noBreak"
                  movel(spat_S_pick_p, a=1.2, v=0.25)
                  # begin: URCap Program Node
                  #   Source: Robotiq_Grippers, 3.17.0.105337, Robotiq Inc.
                  #   Type: Gripper
                  $ 4544 "Gripper Close (1)" "noBreak"
                  if not(gripper_connected[0]):
                    popup("Gripper 1 must be connected to run this program.", "No connection", False, True, True)
                  end
                  if not(rq_is_gripper_activated("1")):
                    popup("Gripper 1 is not activated. Go to Installation tab > Gripper to activate it and run the program again.", "Not activated", False, True, True)
                  end
                  rq_set_pos_spd_for(255, 0, 77, "1")
                  rq_wait_pos_spe_for_request(255, 0, 77, "1")
                  rq_go_to("1")
                  rq_wait("1")
                  # end: URCap Program Node
                  $ 4545 "spat_S_up" "noBreak"
                  movel(spat_S_up_p, a=1.2, v=0.25)
                  $ 4546 "Spatula_otw" "noBreak"
                  movel(Spatula_otw_p, a=1.2, v=0.25)
                  $ 4547 "switch_spat_S≔ False " "noBreak"
                  global switch_spat_S=  False
                  $ 4548 "correction_reset()" "noBreak"
                  correction_reset()
                else:
                  $ 4549 "ElseIf spatula≟'spatula_flat_S'  and switch_spat_F_S ≟ True " "noBreak"
                  if (spatula == "spatula_flat_S"   and  switch_spat_F_S  ==   True  ):
                    $ 4550 "MoveL" "noBreak"
                    $ 4551 "Spatula_otw" "noBreak"
                    movel(Spatula_otw_p, a=1.2, v=0.25)
                    $ 4552 "spat_flatM_up" "noBreak"
                    movel(spat_flatM_up_p, a=1.2, v=0.25)
                    $ 4553 "spat_flatM_pick" "noBreak"
